(* IEC 61131-3 sources: plc-st-coding-agent/progress/evidence/f14_v6_public_pilot_20261112/jobs/codex_deepseek-v4pro, 32 files *)

(* ---- public-easy-01.candidate_01.st ---- *)
(* ENGINEERING_CONTRACT
Output/Public State | Activation (PUB) | Retention/Hold | Reset/Deactivation (PUB) | Same-Scan Priority | Units/Boundaries
Pump_Motor          | bottleSensor (PUB003) | holds through cleaning | cleaningConfirmButton (PUB004) | stage 0 sensor transition first | BOOL, stages 0..5
Filling_Valve       | cleaningConfirmButton (PUB004) | holds through filling | fillingConfirmButton (PUB005) | current stage only | BOOL
Capping_Machine     | fillingConfirmButton (PUB005) | holds through capping | cappingConfirmButton (PUB006) | current stage only | BOOL
Packing_Machine     | cappingConfirmButton (PUB006) | holds through packing | packingConfirmButton (PUB007) | current stage only | BOOL
Completion_Light    | packingConfirmButton (PUB007) | holds until pickup | finishedButton (PUB008) | stage 5 only | BOOL
Unspecified simultaneous assertions are serialized as one stage transition per scan.
*)
(* CONTRACT_RULES [] *)

FUNCTION_BLOCK AutomatedFillingLine
VAR_INPUT
    bottleSensor : BOOL;
    cleaningConfirmButton : BOOL;
    fillingConfirmButton : BOOL;
    cappingConfirmButton : BOOL;
    packingConfirmButton : BOOL;
    finishedButton : BOOL;
END_VAR
VAR_OUTPUT
    Pump_Motor : BOOL;
    Filling_Valve : BOOL;
    Capping_Machine : BOOL;
    Packing_Machine : BOOL;
    Completion_Light : BOOL;
END_VAR
VAR
    tmp_Stage : INT := 0;
END_VAR

CASE tmp_Stage OF
    0:
        IF bottleSensor THEN
            tmp_Stage := 1;
        END_IF;
    1:
        IF cleaningConfirmButton THEN
            tmp_Stage := 2;
        END_IF;
    2:
        IF fillingConfirmButton THEN
            tmp_Stage := 3;
        END_IF;
    3:
        IF cappingConfirmButton THEN
            tmp_Stage := 4;
        END_IF;
    4:
        IF packingConfirmButton THEN
            tmp_Stage := 5;
        END_IF;
    5:
        IF finishedButton THEN
            tmp_Stage := 0;
        END_IF;
END_CASE;

CASE tmp_Stage OF
    0:
        Pump_Motor := FALSE;
        Filling_Valve := FALSE;
        Capping_Machine := FALSE;
        Packing_Machine := FALSE;
        Completion_Light := FALSE;
    1:
        Pump_Motor := TRUE;
        Filling_Valve := FALSE;
        Capping_Machine := FALSE;
        Packing_Machine := FALSE;
        Completion_Light := FALSE;
    2:
        Pump_Motor := FALSE;
        Filling_Valve := TRUE;
        Capping_Machine := FALSE;
        Packing_Machine := FALSE;
        Completion_Light := FALSE;
    3:
        Pump_Motor := FALSE;
        Filling_Valve := FALSE;
        Capping_Machine := TRUE;
        Packing_Machine := FALSE;
        Completion_Light := FALSE;
    4:
        Pump_Motor := FALSE;
        Filling_Valve := FALSE;
        Capping_Machine := FALSE;
        Packing_Machine := TRUE;
        Completion_Light := FALSE;
    5:
        Pump_Motor := FALSE;
        Filling_Valve := FALSE;
        Capping_Machine := FALSE;
        Packing_Machine := FALSE;
        Completion_Light := TRUE;
END_CASE;

END_FUNCTION_BLOCK

(* ---- public-easy-01.candidate_02.st ---- *)
(* ENGINEERING_CONTRACT
Output/Public State | Activation (PUB) | Retention/Hold | Reset/Deactivation (PUB) | Same-Scan Priority | Units/Boundaries
Pump_Motor          | bottleSensor (PUB003) | holds through entire production cycle | finishedButton (PUB008) | stage 0 sensor transition first | BOOL, stages 0..5
Filling_Valve       | cleaningConfirmButton (PUB004) | holds through filling | fillingConfirmButton (PUB005) | current stage only | BOOL
Capping_Machine     | fillingConfirmButton (PUB005) | holds through capping | cappingConfirmButton (PUB006) | current stage only | BOOL
Packing_Machine     | cappingConfirmButton (PUB006) | holds through packing | packingConfirmButton (PUB007) | current stage only | BOOL
Completion_Light    | packingConfirmButton (PUB007) | holds until pickup | finishedButton (PUB008) | stage 5 only | BOOL
Unspecified simultaneous assertions are serialized as one stage transition per scan.
*)
(* CONTRACT_RULES [] *)

FUNCTION_BLOCK AutomatedFillingLine
VAR_INPUT
    bottleSensor : BOOL;
    cleaningConfirmButton : BOOL;
    fillingConfirmButton : BOOL;
    cappingConfirmButton : BOOL;
    packingConfirmButton : BOOL;
    finishedButton : BOOL;
END_VAR
VAR_OUTPUT
    Pump_Motor : BOOL;
    Filling_Valve : BOOL;
    Capping_Machine : BOOL;
    Packing_Machine : BOOL;
    Completion_Light : BOOL;
END_VAR
VAR
    tmp_Stage : INT := 0;
END_VAR

CASE tmp_Stage OF
    0:
        IF bottleSensor THEN
            tmp_Stage := 1;
        END_IF;
    1:
        IF cleaningConfirmButton THEN
            tmp_Stage := 2;
        END_IF;
    2:
        IF fillingConfirmButton THEN
            tmp_Stage := 3;
        END_IF;
    3:
        IF cappingConfirmButton THEN
            tmp_Stage := 4;
        END_IF;
    4:
        IF packingConfirmButton THEN
            tmp_Stage := 5;
        END_IF;
    5:
        IF finishedButton THEN
            tmp_Stage := 0;
        END_IF;
END_CASE;

CASE tmp_Stage OF
    0:
        Pump_Motor := FALSE;
        Filling_Valve := FALSE;
        Capping_Machine := FALSE;
        Packing_Machine := FALSE;
        Completion_Light := FALSE;
    1:
        Pump_Motor := TRUE;
        Filling_Valve := FALSE;
        Capping_Machine := FALSE;
        Packing_Machine := FALSE;
        Completion_Light := FALSE;
    2:
        Pump_Motor := TRUE;
        Filling_Valve := TRUE;
        Capping_Machine := FALSE;
        Packing_Machine := FALSE;
        Completion_Light := FALSE;
    3:
        Pump_Motor := TRUE;
        Filling_Valve := FALSE;
        Capping_Machine := TRUE;
        Packing_Machine := FALSE;
        Completion_Light := FALSE;
    4:
        Pump_Motor := TRUE;
        Filling_Valve := FALSE;
        Capping_Machine := FALSE;
        Packing_Machine := TRUE;
        Completion_Light := FALSE;
    5:
        Pump_Motor := TRUE;
        Filling_Valve := FALSE;
        Capping_Machine := FALSE;
        Packing_Machine := FALSE;
        Completion_Light := TRUE;
END_CASE;

END_FUNCTION_BLOCK

(* ---- public-easy-01.candidate_03.st ---- *)
(* ENGINEERING_CONTRACT
Output/Public State | Activation (PUB) | Retention/Hold | Reset/Deactivation (PUB) | Same-Scan Priority | Units/Boundaries
Pump_Motor          | bottleSensor (PUB003)         | latched after set through cycle | finishedButton (PUB008) | finishedButton reset wins; then set inputs latch | BOOL
Filling_Valve       | cleaningConfirmButton (PUB004) | latched after set through cycle | finishedButton (PUB008) | finishedButton reset wins; then set inputs latch | BOOL
Capping_Machine     | fillingConfirmButton (PUB005)  | latched after set through cycle | finishedButton (PUB008) | finishedButton reset wins; then set inputs latch | BOOL
Packing_Machine     | cappingConfirmButton (PUB006)  | latched after set through cycle | finishedButton (PUB008) | finishedButton reset wins; then set inputs latch | BOOL
Completion_Light    | packingConfirmButton (PUB007)  | latched after set until pickup | finishedButton (PUB008) | finishedButton reset wins; then set inputs latch | BOOL
All BOOL outputs; no step-enable interlock is applied beyond the specified triggers and finished reset.
*)

(* CONTRACT_RULES [
{"kind":"hold_until_reset","output":"Pump_Motor","set_input":"bottleSensor","reset_input":"finishedButton"},
{"kind":"hold_until_reset","output":"Filling_Valve","set_input":"cleaningConfirmButton","reset_input":"finishedButton"},
{"kind":"hold_until_reset","output":"Capping_Machine","set_input":"fillingConfirmButton","reset_input":"finishedButton"},
{"kind":"hold_until_reset","output":"Packing_Machine","set_input":"cappingConfirmButton","reset_input":"finishedButton"},
{"kind":"hold_until_reset","output":"Completion_Light","set_input":"packingConfirmButton","reset_input":"finishedButton"}
] *)

FUNCTION_BLOCK AutomatedFillingLine
VAR_INPUT
    bottleSensor : BOOL;
    cleaningConfirmButton : BOOL;
    fillingConfirmButton : BOOL;
    cappingConfirmButton : BOOL;
    packingConfirmButton : BOOL;
    finishedButton : BOOL;
END_VAR
VAR_OUTPUT
    Pump_Motor : BOOL;
    Filling_Valve : BOOL;
    Capping_Machine : BOOL;
    Packing_Machine : BOOL;
    Completion_Light : BOOL;
END_VAR

IF finishedButton THEN
    Pump_Motor := FALSE;
    Filling_Valve := FALSE;
    Capping_Machine := FALSE;
    Packing_Machine := FALSE;
    Completion_Light := FALSE;
ELSE
    IF bottleSensor THEN
        Pump_Motor := TRUE;
    END_IF;

    IF cleaningConfirmButton THEN
        Filling_Valve := TRUE;
    END_IF;

    IF fillingConfirmButton THEN
        Capping_Machine := TRUE;
    END_IF;

    IF cappingConfirmButton THEN
        Packing_Machine := TRUE;
    END_IF;

    IF packingConfirmButton THEN
        Completion_Light := TRUE;
    END_IF;
END_IF;

END_FUNCTION_BLOCK

(* ---- public-easy-01.candidate_04.st ---- *)
(* ENGINEERING_CONTRACT
Output/Public State | Activation (PUB) | Retention/Hold | Reset/Deactivation | Same-Scan Priority | Units/Boundaries
Pump_Motor | bottleSensor (PUB003) | latched after cycle start | finishedButton (PUB008) | finished reset wins | BOOL
Filling_Valve | cleaningConfirmButton AND Pump_Motor (PUB004) | latched after start | finishedButton (PUB008) | finished reset wins | BOOL
Capping_Machine | fillingConfirmButton AND Filling_Valve (PUB005) | latched after start | finishedButton (PUB008) | finished reset wins | BOOL
Packing_Machine | cappingConfirmButton AND Capping_Machine (PUB006) | latched after start | finishedButton (PUB008) | finished reset wins | BOOL
Completion_Light | packingConfirmButton AND Packing_Machine (PUB007) | latched until pickup | finishedButton (PUB008) | finished reset wins | BOOL
*)

(* CONTRACT_RULES [
 {"kind":"hold_until_reset","output":"Pump_Motor","set_input":"bottleSensor","reset_input":"finishedButton"}
] *)

FUNCTION_BLOCK AutomatedFillingLine
VAR_INPUT
    bottleSensor : BOOL;
    cleaningConfirmButton : BOOL;
    fillingConfirmButton : BOOL;
    cappingConfirmButton : BOOL;
    packingConfirmButton : BOOL;
    finishedButton : BOOL;
END_VAR
VAR_OUTPUT
    Pump_Motor : BOOL;
    Filling_Valve : BOOL;
    Capping_Machine : BOOL;
    Packing_Machine : BOOL;
    Completion_Light : BOOL;
END_VAR

IF finishedButton THEN
    Pump_Motor := FALSE;
    Filling_Valve := FALSE;
    Capping_Machine := FALSE;
    Packing_Machine := FALSE;
    Completion_Light := FALSE;
ELSE
    IF bottleSensor THEN
        Pump_Motor := TRUE;
    END_IF;

    IF cleaningConfirmButton AND Pump_Motor THEN
        Filling_Valve := TRUE;
    END_IF;

    IF fillingConfirmButton AND Filling_Valve THEN
        Capping_Machine := TRUE;
    END_IF;

    IF cappingConfirmButton AND Capping_Machine THEN
        Packing_Machine := TRUE;
    END_IF;

    IF packingConfirmButton AND Packing_Machine THEN
        Completion_Light := TRUE;
    END_IF;
END_IF;

END_FUNCTION_BLOCK

(* ---- public-easy-01.raw_candidate_01.st ---- *)
(* ENGINEERING_CONTRACT
Output/Public State | Activation (PUB) | Retention/Hold | Reset/Deactivation (PUB) | Same-Scan Priority | Units/Boundaries
Pump_Motor          | bottleSensor (PUB003) | holds through cleaning | cleaningConfirmButton (PUB004) | stage 0 sensor transition first | BOOL, stages 0..5
Filling_Valve       | cleaningConfirmButton (PUB004) | holds through filling | fillingConfirmButton (PUB005) | current stage only | BOOL
Capping_Machine     | fillingConfirmButton (PUB005) | holds through capping | cappingConfirmButton (PUB006) | current stage only | BOOL
Packing_Machine     | cappingConfirmButton (PUB006) | holds through packing | packingConfirmButton (PUB007) | current stage only | BOOL
Completion_Light    | packingConfirmButton (PUB007) | holds until pickup | finishedButton (PUB008) | stage 5 only | BOOL
Unspecified simultaneous assertions are serialized as one stage transition per scan.
*)
(* CONTRACT_RULES [] *)

FUNCTION_BLOCK AutomatedFillingLine
VAR_INPUT
    bottleSensor : BOOL;
    cleaningConfirmButton : BOOL;
    fillingConfirmButton : BOOL;
    cappingConfirmButton : BOOL;
    packingConfirmButton : BOOL;
    finishedButton : BOOL;
END_VAR
VAR_OUTPUT
    Pump_Motor : BOOL;
    Filling_Valve : BOOL;
    Capping_Machine : BOOL;
    Packing_Machine : BOOL;
    Completion_Light : BOOL;
END_VAR
VAR
    tmp_Stage : INT := 0;
END_VAR

CASE tmp_Stage OF
    0:
        IF bottleSensor THEN
            tmp_Stage := 1;
        END_IF;
    1:
        IF cleaningConfirmButton THEN
            tmp_Stage := 2;
        END_IF;
    2:
        IF fillingConfirmButton THEN
            tmp_Stage := 3;
        END_IF;
    3:
        IF cappingConfirmButton THEN
            tmp_Stage := 4;
        END_IF;
    4:
        IF packingConfirmButton THEN
            tmp_Stage := 5;
        END_IF;
    5:
        IF finishedButton THEN
            tmp_Stage := 0;
        END_IF;
END_CASE;

CASE tmp_Stage OF
    0:
        Pump_Motor := FALSE;
        Filling_Valve := FALSE;
        Capping_Machine := FALSE;
        Packing_Machine := FALSE;
        Completion_Light := FALSE;
    1:
        Pump_Motor := TRUE;
        Filling_Valve := FALSE;
        Capping_Machine := FALSE;
        Packing_Machine := FALSE;
        Completion_Light := FALSE;
    2:
        Pump_Motor := FALSE;
        Filling_Valve := TRUE;
        Capping_Machine := FALSE;
        Packing_Machine := FALSE;
        Completion_Light := FALSE;
    3:
        Pump_Motor := FALSE;
        Filling_Valve := FALSE;
        Capping_Machine := TRUE;
        Packing_Machine := FALSE;
        Completion_Light := FALSE;
    4:
        Pump_Motor := FALSE;
        Filling_Valve := FALSE;
        Capping_Machine := FALSE;
        Packing_Machine := TRUE;
        Completion_Light := FALSE;
    5:
        Pump_Motor := FALSE;
        Filling_Valve := FALSE;
        Capping_Machine := FALSE;
        Packing_Machine := FALSE;
        Completion_Light := TRUE;
END_CASE;

END_FUNCTION_BLOCK

(* ---- public-easy-01.raw_candidate_02.st ---- *)
(* ENGINEERING_CONTRACT
Output/Public State | Activation (PUB) | Retention/Hold | Reset/Deactivation (PUB) | Same-Scan Priority | Units/Boundaries
Pump_Motor          | bottleSensor (PUB003) | holds through entire production cycle | finishedButton (PUB008) | stage 0 sensor transition first | BOOL, stages 0..5
Filling_Valve       | cleaningConfirmButton (PUB004) | holds through filling | fillingConfirmButton (PUB005) | current stage only | BOOL
Capping_Machine     | fillingConfirmButton (PUB005) | holds through capping | cappingConfirmButton (PUB006) | current stage only | BOOL
Packing_Machine     | cappingConfirmButton (PUB006) | holds through packing | packingConfirmButton (PUB007) | current stage only | BOOL
Completion_Light    | packingConfirmButton (PUB007) | holds until pickup | finishedButton (PUB008) | stage 5 only | BOOL
Unspecified simultaneous assertions are serialized as one stage transition per scan.
*)
(* CONTRACT_RULES [] *)

FUNCTION_BLOCK AutomatedFillingLine
VAR_INPUT
    bottleSensor : BOOL;
    cleaningConfirmButton : BOOL;
    fillingConfirmButton : BOOL;
    cappingConfirmButton : BOOL;
    packingConfirmButton : BOOL;
    finishedButton : BOOL;
END_VAR
VAR_OUTPUT
    Pump_Motor : BOOL;
    Filling_Valve : BOOL;
    Capping_Machine : BOOL;
    Packing_Machine : BOOL;
    Completion_Light : BOOL;
END_VAR
VAR
    tmp_Stage : INT := 0;
END_VAR

CASE tmp_Stage OF
    0:
        IF bottleSensor THEN
            tmp_Stage := 1;
        END_IF;
    1:
        IF cleaningConfirmButton THEN
            tmp_Stage := 2;
        END_IF;
    2:
        IF fillingConfirmButton THEN
            tmp_Stage := 3;
        END_IF;
    3:
        IF cappingConfirmButton THEN
            tmp_Stage := 4;
        END_IF;
    4:
        IF packingConfirmButton THEN
            tmp_Stage := 5;
        END_IF;
    5:
        IF finishedButton THEN
            tmp_Stage := 0;
        END_IF;
END_CASE;

CASE tmp_Stage OF
    0:
        Pump_Motor := FALSE;
        Filling_Valve := FALSE;
        Capping_Machine := FALSE;
        Packing_Machine := FALSE;
        Completion_Light := FALSE;
    1:
        Pump_Motor := TRUE;
        Filling_Valve := FALSE;
        Capping_Machine := FALSE;
        Packing_Machine := FALSE;
        Completion_Light := FALSE;
    2:
        Pump_Motor := TRUE;
        Filling_Valve := TRUE;
        Capping_Machine := FALSE;
        Packing_Machine := FALSE;
        Completion_Light := FALSE;
    3:
        Pump_Motor := TRUE;
        Filling_Valve := FALSE;
        Capping_Machine := TRUE;
        Packing_Machine := FALSE;
        Completion_Light := FALSE;
    4:
        Pump_Motor := TRUE;
        Filling_Valve := FALSE;
        Capping_Machine := FALSE;
        Packing_Machine := TRUE;
        Completion_Light := FALSE;
    5:
        Pump_Motor := TRUE;
        Filling_Valve := FALSE;
        Capping_Machine := FALSE;
        Packing_Machine := FALSE;
        Completion_Light := TRUE;
END_CASE;

END_FUNCTION_BLOCK

(* ---- public-easy-01.raw_candidate_03.st ---- *)
(* ENGINEERING_CONTRACT
Output/Public State | Activation (PUB) | Retention/Hold | Reset/Deactivation (PUB) | Same-Scan Priority | Units/Boundaries
Pump_Motor          | bottleSensor (PUB003)         | latched after set through cycle | finishedButton (PUB008) | finishedButton reset wins; then set inputs latch | BOOL
Filling_Valve       | cleaningConfirmButton (PUB004) | latched after set through cycle | finishedButton (PUB008) | finishedButton reset wins; then set inputs latch | BOOL
Capping_Machine     | fillingConfirmButton (PUB005)  | latched after set through cycle | finishedButton (PUB008) | finishedButton reset wins; then set inputs latch | BOOL
Packing_Machine     | cappingConfirmButton (PUB006)  | latched after set through cycle | finishedButton (PUB008) | finishedButton reset wins; then set inputs latch | BOOL
Completion_Light    | packingConfirmButton (PUB007)  | latched after set until pickup | finishedButton (PUB008) | finishedButton reset wins; then set inputs latch | BOOL
All BOOL outputs; no step-enable interlock is applied beyond the specified triggers and finished reset.
*)

(* CONTRACT_RULES [
{"kind":"hold_until_reset","output":"Pump_Motor","set_input":"bottleSensor","reset_input":"finishedButton"},
{"kind":"hold_until_reset","output":"Filling_Valve","set_input":"cleaningConfirmButton","reset_input":"finishedButton"},
{"kind":"hold_until_reset","output":"Capping_Machine","set_input":"fillingConfirmButton","reset_input":"finishedButton"},
{"kind":"hold_until_reset","output":"Packing_Machine","set_input":"cappingConfirmButton","reset_input":"finishedButton"},
{"kind":"hold_until_reset","output":"Completion_Light","set_input":"packingConfirmButton","reset_input":"finishedButton"}
] *)

FUNCTION_BLOCK AutomatedFillingLine
VAR_INPUT
    bottleSensor : BOOL;
    cleaningConfirmButton : BOOL;
    fillingConfirmButton : BOOL;
    cappingConfirmButton : BOOL;
    packingConfirmButton : BOOL;
    finishedButton : BOOL;
END_VAR
VAR_OUTPUT
    Pump_Motor : BOOL;
    Filling_Valve : BOOL;
    Capping_Machine : BOOL;
    Packing_Machine : BOOL;
    Completion_Light : BOOL;
END_VAR

IF finishedButton THEN
    Pump_Motor := FALSE;
    Filling_Valve := FALSE;
    Capping_Machine := FALSE;
    Packing_Machine := FALSE;
    Completion_Light := FALSE;
ELSE
    IF bottleSensor THEN
        Pump_Motor := TRUE;
    END_IF;

    IF cleaningConfirmButton THEN
        Filling_Valve := TRUE;
    END_IF;

    IF fillingConfirmButton THEN
        Capping_Machine := TRUE;
    END_IF;

    IF cappingConfirmButton THEN
        Packing_Machine := TRUE;
    END_IF;

    IF packingConfirmButton THEN
        Completion_Light := TRUE;
    END_IF;
END_IF;

END_FUNCTION_BLOCK

(* ---- public-easy-01.raw_candidate_04.st ---- *)
(* ENGINEERING_CONTRACT
Output/Public State | Activation (PUB) | Retention/Hold | Reset/Deactivation | Same-Scan Priority | Units/Boundaries
Pump_Motor | bottleSensor (PUB003) | latched after cycle start | finishedButton (PUB008) | finished reset wins | BOOL
Filling_Valve | cleaningConfirmButton AND Pump_Motor (PUB004) | latched after start | finishedButton (PUB008) | finished reset wins | BOOL
Capping_Machine | fillingConfirmButton AND Filling_Valve (PUB005) | latched after start | finishedButton (PUB008) | finished reset wins | BOOL
Packing_Machine | cappingConfirmButton AND Capping_Machine (PUB006) | latched after start | finishedButton (PUB008) | finished reset wins | BOOL
Completion_Light | packingConfirmButton AND Packing_Machine (PUB007) | latched until pickup | finishedButton (PUB008) | finished reset wins | BOOL
*)

(* CONTRACT_RULES [
 {"kind":"hold_until_reset","output":"Pump_Motor","set_input":"bottleSensor","reset_input":"finishedButton"}
] *)

FUNCTION_BLOCK AutomatedFillingLine
VAR_INPUT
    bottleSensor : BOOL;
    cleaningConfirmButton : BOOL;
    fillingConfirmButton : BOOL;
    cappingConfirmButton : BOOL;
    packingConfirmButton : BOOL;
    finishedButton : BOOL;
END_VAR
VAR_OUTPUT
    Pump_Motor : BOOL;
    Filling_Valve : BOOL;
    Capping_Machine : BOOL;
    Packing_Machine : BOOL;
    Completion_Light : BOOL;
END_VAR

IF finishedButton THEN
    Pump_Motor := FALSE;
    Filling_Valve := FALSE;
    Capping_Machine := FALSE;
    Packing_Machine := FALSE;
    Completion_Light := FALSE;
ELSE
    IF bottleSensor THEN
        Pump_Motor := TRUE;
    END_IF;

    IF cleaningConfirmButton AND Pump_Motor THEN
        Filling_Valve := TRUE;
    END_IF;

    IF fillingConfirmButton AND Filling_Valve THEN
        Capping_Machine := TRUE;
    END_IF;

    IF cappingConfirmButton AND Capping_Machine THEN
        Packing_Machine := TRUE;
    END_IF;

    IF packingConfirmButton AND Packing_Machine THEN
        Completion_Light := TRUE;
    END_IF;
END_IF;

END_FUNCTION_BLOCK

(* ---- public-easy-04.candidate_01.st ---- *)
(*
ENGINEERING_CONTRACT
- VFD_RUN: active iff PASTE_E_STOP_NC AND viscosity_condition; no retention; immediate off on raw FALSE or E_STOP FALSE; PUB003.
- viscosity_condition: becomes TRUE when VISCOSITY_OK TRUE for >= DebounceTime; raw FALSE invalidates immediately; E_STOP clears only incomplete debounce; PUB002/PUB003.
- PUMP_RUNTIME_ACC: adds TIME_TO_LTIME(CycleTime) only when final VFD_RUN TRUE; preserved while stopped; starts at zero; PUB004/PUB006.
- PUMP_MAINT_DUE: TRUE when PUMP_RUNTIME_ACC >= TIME_TO_LTIME(T#500H); informational, no run/permissive effect; PUB005.
- units: DebounceTime/CycleTime TIME ms; accumulated value LTIME ns.
- priority: raw viscosity FALSE and E_STOP FALSE are resolved before same-scan runtime accumulation.
*)
(* CONTRACT_RULES [] *)

FUNCTION_BLOCK JamPumpControl
VAR_INPUT
    VISCOSITY_OK : BOOL;
    PASTE_E_STOP_NC : BOOL;
    DebounceTime : TIME;
    CycleTime : TIME;
END_VAR
VAR_OUTPUT
    VFD_RUN : BOOL;
    PUMP_MAINT_DUE : BOOL;
    PUMP_RUNTIME_ACC : LTIME;
END_VAR
VAR
    local_debounce_elapsed : LTIME := LTIME#0S;
    local_viscosity_condition : BOOL := FALSE;
    local_runtime_accumulator : LTIME := LTIME#0S;
END_VAR

IF VISCOSITY_OK THEN
    IF PASTE_E_STOP_NC THEN
        IF CycleTime > T#0MS THEN
            IF local_debounce_elapsed < TIME_TO_LTIME(DebounceTime) THEN
                local_debounce_elapsed := local_debounce_elapsed + TIME_TO_LTIME(CycleTime);
                IF local_debounce_elapsed > TIME_TO_LTIME(DebounceTime) THEN
                    local_debounce_elapsed := TIME_TO_LTIME(DebounceTime);
                END_IF;
            END_IF;
        END_IF;
    ELSE
        IF local_debounce_elapsed < TIME_TO_LTIME(DebounceTime) THEN
            local_debounce_elapsed := LTIME#0S;
            local_viscosity_condition := FALSE;
        END_IF;
    END_IF;
    local_viscosity_condition := local_debounce_elapsed >= TIME_TO_LTIME(DebounceTime);
ELSE
    local_debounce_elapsed := LTIME#0S;
    local_viscosity_condition := FALSE;
END_IF;

VFD_RUN := PASTE_E_STOP_NC AND local_viscosity_condition;

IF VFD_RUN THEN
    IF CycleTime > T#0MS THEN
        local_runtime_accumulator := local_runtime_accumulator + TIME_TO_LTIME(CycleTime);
    END_IF;
END_IF;

PUMP_RUNTIME_ACC := local_runtime_accumulator;
PUMP_MAINT_DUE := local_runtime_accumulator >= TIME_TO_LTIME(T#500H);

END_FUNCTION_BLOCK

(* ---- public-easy-04.raw_candidate_01.st ---- *)
(*
ENGINEERING_CONTRACT
- VFD_RUN: active iff PASTE_E_STOP_NC AND viscosity_condition; no retention; immediate off on raw FALSE or E_STOP FALSE; PUB003.
- viscosity_condition: becomes TRUE when VISCOSITY_OK TRUE for >= DebounceTime; raw FALSE invalidates immediately; E_STOP clears only incomplete debounce; PUB002/PUB003.
- PUMP_RUNTIME_ACC: adds TIME_TO_LTIME(CycleTime) only when final VFD_RUN TRUE; preserved while stopped; starts at zero; PUB004/PUB006.
- PUMP_MAINT_DUE: TRUE when PUMP_RUNTIME_ACC >= TIME_TO_LTIME(T#500H); informational, no run/permissive effect; PUB005.
- units: DebounceTime/CycleTime TIME ms; accumulated value LTIME ns.
- priority: raw viscosity FALSE and E_STOP FALSE are resolved before same-scan runtime accumulation.
*)
(* CONTRACT_RULES [] *)

FUNCTION_BLOCK JamPumpControl
VAR_INPUT
    VISCOSITY_OK : BOOL;
    PASTE_E_STOP_NC : BOOL;
    DebounceTime : TIME;
    CycleTime : TIME;
END_VAR
VAR_OUTPUT
    VFD_RUN : BOOL;
    PUMP_MAINT_DUE : BOOL;
    PUMP_RUNTIME_ACC : LTIME;
END_VAR
VAR
    local_debounce_elapsed : LTIME := LTIME#0S;
    local_viscosity_condition : BOOL := FALSE;
    local_runtime_accumulator : LTIME := LTIME#0S;
END_VAR

IF VISCOSITY_OK THEN
    IF PASTE_E_STOP_NC THEN
        IF CycleTime > T#0MS THEN
            IF local_debounce_elapsed < TIME_TO_LTIME(DebounceTime) THEN
                local_debounce_elapsed := local_debounce_elapsed + TIME_TO_LTIME(CycleTime);
                IF local_debounce_elapsed > TIME_TO_LTIME(DebounceTime) THEN
                    local_debounce_elapsed := TIME_TO_LTIME(DebounceTime);
                END_IF;
            END_IF;
        END_IF;
    ELSE
        IF local_debounce_elapsed < TIME_TO_LTIME(DebounceTime) THEN
            local_debounce_elapsed := LTIME#0S;
            local_viscosity_condition := FALSE;
        END_IF;
    END_IF;
    local_viscosity_condition := local_debounce_elapsed >= TIME_TO_LTIME(DebounceTime);
ELSE
    local_debounce_elapsed := LTIME#0S;
    local_viscosity_condition := FALSE;
END_IF;

VFD_RUN := PASTE_E_STOP_NC AND local_viscosity_condition;

IF VFD_RUN THEN
    IF CycleTime > T#0MS THEN
        local_runtime_accumulator := local_runtime_accumulator + TIME_TO_LTIME(CycleTime);
    END_IF;
END_IF;

PUMP_RUNTIME_ACC := local_runtime_accumulator;
PUMP_MAINT_DUE := local_runtime_accumulator >= TIME_TO_LTIME(T#500H);

END_FUNCTION_BLOCK

(* ---- public-hard-03.candidate_01.st ---- *)
TYPE ST_Recipe :
STRUCT
    recipeID : INT;
    ingredientType : INT;
    ingredientRatio : REAL;
    productionTemperature : REAL;
END_STRUCT
END_TYPE;

FUNCTION_BLOCK FB_RecipeManager
VAR_INPUT
    addRecipe : BOOL;
    deleteRecipe : BOOL;
    modifyRecipe : BOOL;
    queryRecipe : BOOL;
    recipeIn : ST_Recipe;
END_VAR
VAR_OUTPUT
    recipeAdded : BOOL;
    recipeDeleted : BOOL;
    recipeModified : BOOL;
    recipeQueryResult : ST_Recipe;
    error : BOOL;
    status : WORD;
END_VAR
VAR_IN_OUT
    recipe : ARRAY[1..10] OF ST_Recipe;
END_VAR
VAR
    local_i : INT;
    local_matchIndex : INT;
    local_emptyIndex : INT;
    local_found : BOOL;
    local_emptyFound : BOOL;
    local_activeCommands : INT;
END_VAR

(* ENGINEERING_CONTRACT
  Outputs/database behavior:
  - recipeAdded/recipeDeleted/recipeModified: TRUE only on a successful same-scan command, cleared each scan; no hold.
  - recipeQueryResult: written only on a successful query, cleared at scan start; no retention.
  - error/status: set on command failures per PUB009-PUB012, cleared each scan; no hold.
  - Add order: duplicate=16#8002 before full=16#8003; success fills smallest empty index (PUB010).
  - Delete sets only matching recipeID to 0 (PUB011); modify replaces matching slot (PUB012).
  - recipeID 0 is an empty slot marker. Query/delete/modify of ID 0 returns command-specific failure.
  - Multiple simultaneous commands are unsupported: error=TRUE, status=16#80FF, database unchanged.
  - Bounds: array[1..10], IDs INT, ratios/temperatures REAL (PUB008).
*)

(* CONTRACT_RULES [] *)

recipeAdded := FALSE;
recipeDeleted := FALSE;
recipeModified := FALSE;
recipeQueryResult.recipeID := 0;
recipeQueryResult.ingredientType := 0;
recipeQueryResult.ingredientRatio := 0.0;
recipeQueryResult.productionTemperature := 0.0;
error := FALSE;
status := 16#0000;

local_activeCommands := BOOL_TO_INT(addRecipe) + BOOL_TO_INT(deleteRecipe) + BOOL_TO_INT(modifyRecipe) + BOOL_TO_INT(queryRecipe);

IF local_activeCommands > 1 THEN
    error := TRUE;
    status := 16#80FF;
    RETURN;
END_IF;

IF queryRecipe THEN
    local_found := FALSE;
    local_matchIndex := 0;

    IF recipeIn.recipeID <> 0 THEN
        FOR local_i := 1 TO 10 BY 1 DO
            IF (NOT local_found) AND (recipe[local_i].recipeID = recipeIn.recipeID) THEN
                local_matchIndex := local_i;
                local_found := TRUE;
            END_IF;
        END_FOR;
    END_IF;

    IF local_found THEN
        recipeQueryResult := recipe[local_matchIndex];
        error := FALSE;
        status := 16#0000;
    ELSE
        error := TRUE;
        status := 16#8001;
    END_IF;

ELSIF addRecipe THEN
    local_found := FALSE;
    local_emptyFound := FALSE;
    local_emptyIndex := 0;

    FOR local_i := 1 TO 10 BY 1 DO
        IF recipe[local_i].recipeID = recipeIn.recipeID THEN
            local_found := TRUE;
        END_IF;

        IF (NOT local_emptyFound) AND (recipe[local_i].recipeID = 0) THEN
            local_emptyIndex := local_i;
            local_emptyFound := TRUE;
        END_IF;
    END_FOR;

    IF local_found THEN
        error := TRUE;
        status := 16#8002;
    ELSIF NOT local_emptyFound THEN
        error := TRUE;
        status := 16#8003;
    ELSE
        recipe[local_emptyIndex] := recipeIn;
        recipeAdded := TRUE;
        error := FALSE;
        status := 16#0000;
    END_IF;

ELSIF deleteRecipe THEN
    local_found := FALSE;
    local_matchIndex := 0;

    IF recipeIn.recipeID <> 0 THEN
        FOR local_i := 1 TO 10 BY 1 DO
            IF (NOT local_found) AND (recipe[local_i].recipeID = recipeIn.recipeID) THEN
                local_matchIndex := local_i;
                local_found := TRUE;
            END_IF;
        END_FOR;
    END_IF;

    IF local_found THEN
        recipe[local_matchIndex].recipeID := 0;
        recipeDeleted := TRUE;
        error := FALSE;
        status := 16#0000;
    ELSE
        error := TRUE;
        status := 16#8004;
    END_IF;

ELSIF modifyRecipe THEN
    local_found := FALSE;
    local_matchIndex := 0;

    IF recipeIn.recipeID <> 0 THEN
        FOR local_i := 1 TO 10 BY 1 DO
            IF (NOT local_found) AND (recipe[local_i].recipeID = recipeIn.recipeID) THEN
                local_matchIndex := local_i;
                local_found := TRUE;
            END_IF;
        END_FOR;
    END_IF;

    IF local_found THEN
        recipe[local_matchIndex] := recipeIn;
        recipeModified := TRUE;
        error := FALSE;
        status := 16#0000;
    ELSE
        error := TRUE;
        status := 16#8005;
    END_IF;
END_IF;
END_FUNCTION_BLOCK

(* ---- public-hard-03.candidate_02.st ---- *)
TYPE ST_Recipe :
STRUCT
    recipeID : INT;
    ingredientType : INT;
    ingredientRatio : REAL;
    productionTemperature : REAL;
END_STRUCT
END_TYPE;

FUNCTION_BLOCK FB_RecipeManager
VAR_INPUT
    addRecipe : BOOL;
    deleteRecipe : BOOL;
    modifyRecipe : BOOL;
    queryRecipe : BOOL;
    recipeIn : ST_Recipe;
END_VAR
VAR_OUTPUT
    recipeAdded : BOOL;
    recipeDeleted : BOOL;
    recipeModified : BOOL;
    recipeQueryResult : ST_Recipe;
    error : BOOL;
    status : WORD;
END_VAR
VAR_IN_OUT
    recipe : ARRAY[1..10] OF ST_Recipe;
END_VAR
VAR
    local_i : INT;
    local_matchIndex : INT;
    local_emptyIndex : INT;
    local_found : BOOL;
    local_emptyFound : BOOL;
END_VAR

(* ENGINEERING_CONTRACT
  Outputs/database behavior:
  - recipeAdded/recipeDeleted/recipeModified: pulse TRUE only on a successful same-scan command, cleared at scan start.
  - recipeQueryResult: cleared at scan start; rewritten only on a successful query.
  - error/status: set on command failure per PUB009-PUB012, otherwise no error.
  - Add checks duplicate before full, then stores at smallest empty index (PUB010).
  - Delete clears only the matching recipeID (PUB011); modify replaces the matching slot (PUB012).
  - Query ID not found => error=TRUE, status=16#8001 (PUB009).
  - Add duplicate => 16#8002; add full => 16#8003 (PUB010).
  - Delete ID not found => 16#8004 (PUB011); modify ID not found => 16#8005 (PUB012).
  - recipeID 0 denotes an empty slot (PUB008).
  - Simultaneous commands are unspecified by task text; implemented with interface-order priority:
    addRecipe > deleteRecipe > modifyRecipe > queryRecipe. The higher-priority command is executed,
    lower-priority commands are not processed in that scan.
  - Bounds: ARRAY[1..10], INT and REAL data preserved exactly (PUB008).
*)

(* CONTRACT_RULES [] *)

recipeAdded := FALSE;
recipeDeleted := FALSE;
recipeModified := FALSE;
recipeQueryResult.recipeID := 0;
recipeQueryResult.ingredientType := 0;
recipeQueryResult.ingredientRatio := 0.0;
recipeQueryResult.productionTemperature := 0.0;
error := FALSE;
status := 16#0000;

IF addRecipe THEN
    local_found := FALSE;
    local_emptyFound := FALSE;
    local_emptyIndex := 0;

    FOR local_i := 1 TO 10 BY 1 DO
        IF recipe[local_i].recipeID = recipeIn.recipeID THEN
            local_found := TRUE;
        END_IF;

        IF (NOT local_emptyFound) AND (recipe[local_i].recipeID = 0) THEN
            local_emptyIndex := local_i;
            local_emptyFound := TRUE;
        END_IF;
    END_FOR;

    IF local_found THEN
        error := TRUE;
        status := 16#8002;
    ELSIF NOT local_emptyFound THEN
        error := TRUE;
        status := 16#8003;
    ELSE
        recipe[local_emptyIndex] := recipeIn;
        recipeAdded := TRUE;
        error := FALSE;
        status := 16#0000;
    END_IF;

ELSIF deleteRecipe THEN
    local_found := FALSE;
    local_matchIndex := 0;

    IF recipeIn.recipeID <> 0 THEN
        FOR local_i := 1 TO 10 BY 1 DO
            IF (NOT local_found) AND (recipe[local_i].recipeID = recipeIn.recipeID) THEN
                local_matchIndex := local_i;
                local_found := TRUE;
            END_IF;
        END_FOR;
    END_IF;

    IF local_found THEN
        recipe[local_matchIndex].recipeID := 0;
        recipeDeleted := TRUE;
        error := FALSE;
        status := 16#0000;
    ELSE
        error := TRUE;
        status := 16#8004;
    END_IF;

ELSIF modifyRecipe THEN
    local_found := FALSE;
    local_matchIndex := 0;

    IF recipeIn.recipeID <> 0 THEN
        FOR local_i := 1 TO 10 BY 1 DO
            IF (NOT local_found) AND (recipe[local_i].recipeID = recipeIn.recipeID) THEN
                local_matchIndex := local_i;
                local_found := TRUE;
            END_IF;
        END_FOR;
    END_IF;

    IF local_found THEN
        recipe[local_matchIndex] := recipeIn;
        recipeModified := TRUE;
        error := FALSE;
        status := 16#0000;
    ELSE
        error := TRUE;
        status := 16#8005;
    END_IF;

ELSIF queryRecipe THEN
    local_found := FALSE;
    local_matchIndex := 0;

    IF recipeIn.recipeID <> 0 THEN
        FOR local_i := 1 TO 10 BY 1 DO
            IF (NOT local_found) AND (recipe[local_i].recipeID = recipeIn.recipeID) THEN
                local_matchIndex := local_i;
                local_found := TRUE;
            END_IF;
        END_FOR;
    END_IF;

    IF local_found THEN
        recipeQueryResult := recipe[local_matchIndex];
        error := FALSE;
        status := 16#0000;
    ELSE
        error := TRUE;
        status := 16#8001;
    END_IF;
END_IF;
END_FUNCTION_BLOCK

(* ---- public-hard-03.candidate_03.st ---- *)
TYPE ST_Recipe :
STRUCT
    recipeID : INT;
    ingredientType : INT;
    ingredientRatio : REAL;
    productionTemperature : REAL;
END_STRUCT
END_TYPE;

FUNCTION_BLOCK FB_RecipeManager
VAR_INPUT
    addRecipe : BOOL;
    deleteRecipe : BOOL;
    modifyRecipe : BOOL;
    queryRecipe : BOOL;
    recipeIn : ST_Recipe;
END_VAR
VAR_OUTPUT
    recipeAdded : BOOL;
    recipeDeleted : BOOL;
    recipeModified : BOOL;
    recipeQueryResult : ST_Recipe;
    error : BOOL;
    status : WORD;
END_VAR
VAR_IN_OUT
    recipe : ARRAY[1..10] OF ST_Recipe;
END_VAR
VAR
    local_i : INT;
    local_matchIndex : INT;
    local_emptyIndex : INT;
    local_found : BOOL;
    local_emptyFound : BOOL;
END_VAR

(* ENGINEERING_CONTRACT
  Outputs/database behavior:
  - recipeAdded/recipeDeleted/recipeModified: TRUE only on a successful same-scan command, cleared each scan; no hold.
  - recipeQueryResult: written only on a successful query, cleared at scan start; no retention.
  - error/status: set on command failures per PUB009-PUB012, cleared each scan; no hold.
  - Simultaneous commands: addRecipe has priority; then queryRecipe, deleteRecipe, modifyRecipe.
  - Add order: duplicate=16#8002 before full=16#8003; success fills smallest empty index (PUB010).
  - Delete sets only matching recipeID to 0 (PUB011); modify replaces matching slot (PUB012).
  - recipeID 0 is an empty slot marker. Query/delete/modify of ID 0 returns command-specific failure.
  - Bounds: array[1..10], IDs INT, ratios/temperatures REAL (PUB008).
*)

(* CONTRACT_RULES [] *)

recipeAdded := FALSE;
recipeDeleted := FALSE;
recipeModified := FALSE;
recipeQueryResult.recipeID := 0;
recipeQueryResult.ingredientType := 0;
recipeQueryResult.ingredientRatio := 0.0;
recipeQueryResult.productionTemperature := 0.0;
error := FALSE;
status := 16#0000;

IF addRecipe THEN
    local_found := FALSE;
    local_emptyFound := FALSE;
    local_emptyIndex := 0;

    FOR local_i := 1 TO 10 BY 1 DO
        IF recipe[local_i].recipeID = recipeIn.recipeID THEN
            local_found := TRUE;
        END_IF;

        IF (NOT local_emptyFound) AND (recipe[local_i].recipeID = 0) THEN
            local_emptyIndex := local_i;
            local_emptyFound := TRUE;
        END_IF;
    END_FOR;

    IF local_found THEN
        error := TRUE;
        status := 16#8002;
    ELSIF NOT local_emptyFound THEN
        error := TRUE;
        status := 16#8003;
    ELSE
        recipe[local_emptyIndex] := recipeIn;
        recipeAdded := TRUE;
        error := FALSE;
        status := 16#0000;
    END_IF;

ELSIF queryRecipe THEN
    local_found := FALSE;
    local_matchIndex := 0;

    IF recipeIn.recipeID <> 0 THEN
        FOR local_i := 1 TO 10 BY 1 DO
            IF (NOT local_found) AND (recipe[local_i].recipeID = recipeIn.recipeID) THEN
                local_matchIndex := local_i;
                local_found := TRUE;
            END_IF;
        END_FOR;
    END_IF;

    IF local_found THEN
        recipeQueryResult := recipe[local_matchIndex];
        error := FALSE;
        status := 16#0000;
    ELSE
        error := TRUE;
        status := 16#8001;
    END_IF;

ELSIF deleteRecipe THEN
    local_found := FALSE;
    local_matchIndex := 0;

    IF recipeIn.recipeID <> 0 THEN
        FOR local_i := 1 TO 10 BY 1 DO
            IF (NOT local_found) AND (recipe[local_i].recipeID = recipeIn.recipeID) THEN
                local_matchIndex := local_i;
                local_found := TRUE;
            END_IF;
        END_FOR;
    END_IF;

    IF local_found THEN
        recipe[local_matchIndex].recipeID := 0;
        recipeDeleted := TRUE;
        error := FALSE;
        status := 16#0000;
    ELSE
        error := TRUE;
        status := 16#8004;
    END_IF;

ELSIF modifyRecipe THEN
    local_found := FALSE;
    local_matchIndex := 0;

    IF recipeIn.recipeID <> 0 THEN
        FOR local_i := 1 TO 10 BY 1 DO
            IF (NOT local_found) AND (recipe[local_i].recipeID = recipeIn.recipeID) THEN
                local_matchIndex := local_i;
                local_found := TRUE;
            END_IF;
        END_FOR;
    END_IF;

    IF local_found THEN
        recipe[local_matchIndex] := recipeIn;
        recipeModified := TRUE;
        error := FALSE;
        status := 16#0000;
    ELSE
        error := TRUE;
        status := 16#8005;
    END_IF;
END_IF;
END_FUNCTION_BLOCK

(* ---- public-hard-03.candidate_04.st ---- *)
TYPE ST_Recipe :
STRUCT
    recipeID : INT;
    ingredientType : INT;
    ingredientRatio : REAL;
    productionTemperature : REAL;
END_STRUCT
END_TYPE;

FUNCTION_BLOCK FB_RecipeManager
VAR_INPUT
    addRecipe : BOOL;
    deleteRecipe : BOOL;
    modifyRecipe : BOOL;
    queryRecipe : BOOL;
    recipeIn : ST_Recipe;
END_VAR
VAR_OUTPUT
    recipeAdded : BOOL;
    recipeDeleted : BOOL;
    recipeModified : BOOL;
    recipeQueryResult : ST_Recipe;
    error : BOOL;
    status : WORD;
END_VAR
VAR_IN_OUT
    recipe : ARRAY[1..10] OF ST_Recipe;
END_VAR
VAR
    local_i : INT;
    local_matchIndex : INT;
    local_emptyIndex : INT;
    local_found : BOOL;
    local_emptyFound : BOOL;
END_VAR

(* ENGINEERING_CONTRACT
  Outputs/database behavior:
  - recipeAdded/recipeDeleted/recipeModified: TRUE only on a successful same-scan command, cleared each scan; no hold.
  - recipeQueryResult: written only on a successful query, cleared at scan start; no retention.
  - error/status: set on command failures per PUB009-PUB012, cleared each scan; no hold.
  - Add order: duplicate=16#8002 before full=16#8003; success fills smallest empty index (PUB010).
  - Delete sets only matching recipeID to 0 (PUB011); modify replaces matching slot (PUB012).
  - recipeID 0 is an empty slot marker. Query/delete/modify of ID 0 returns command-specific failure.
  - Multiple simultaneous commands are unspecified by PUB. Consistent interpretation: add > delete > modify > query.
  - Bounds: array[1..10], IDs INT, ratios/temperatures REAL (PUB008).
*)

(* CONTRACT_RULES [] *)

recipeAdded := FALSE;
recipeDeleted := FALSE;
recipeModified := FALSE;
recipeQueryResult.recipeID := 0;
recipeQueryResult.ingredientType := 0;
recipeQueryResult.ingredientRatio := 0.0;
recipeQueryResult.productionTemperature := 0.0;
error := FALSE;
status := 16#0000;

IF addRecipe THEN
    local_found := FALSE;
    local_emptyFound := FALSE;
    local_emptyIndex := 0;

    FOR local_i := 1 TO 10 BY 1 DO
        IF recipe[local_i].recipeID = recipeIn.recipeID THEN
            local_found := TRUE;
        END_IF;

        IF (NOT local_emptyFound) AND (recipe[local_i].recipeID = 0) THEN
            local_emptyIndex := local_i;
            local_emptyFound := TRUE;
        END_IF;
    END_FOR;

    IF local_found THEN
        error := TRUE;
        status := 16#8002;
    ELSIF NOT local_emptyFound THEN
        error := TRUE;
        status := 16#8003;
    ELSE
        recipe[local_emptyIndex] := recipeIn;
        recipeAdded := TRUE;
        error := FALSE;
        status := 16#0000;
    END_IF;

ELSIF deleteRecipe THEN
    local_found := FALSE;
    local_matchIndex := 0;

    IF recipeIn.recipeID <> 0 THEN
        FOR local_i := 1 TO 10 BY 1 DO
            IF (NOT local_found) AND (recipe[local_i].recipeID = recipeIn.recipeID) THEN
                local_matchIndex := local_i;
                local_found := TRUE;
            END_IF;
        END_FOR;
    END_IF;

    IF local_found THEN
        recipe[local_matchIndex].recipeID := 0;
        recipeDeleted := TRUE;
        error := FALSE;
        status := 16#0000;
    ELSE
        error := TRUE;
        status := 16#8004;
    END_IF;

ELSIF modifyRecipe THEN
    local_found := FALSE;
    local_matchIndex := 0;

    IF recipeIn.recipeID <> 0 THEN
        FOR local_i := 1 TO 10 BY 1 DO
            IF (NOT local_found) AND (recipe[local_i].recipeID = recipeIn.recipeID) THEN
                local_matchIndex := local_i;
                local_found := TRUE;
            END_IF;
        END_FOR;
    END_IF;

    IF local_found THEN
        recipe[local_matchIndex] := recipeIn;
        recipeModified := TRUE;
        error := FALSE;
        status := 16#0000;
    ELSE
        error := TRUE;
        status := 16#8005;
    END_IF;

ELSIF queryRecipe THEN
    local_found := FALSE;
    local_matchIndex := 0;

    IF recipeIn.recipeID <> 0 THEN
        FOR local_i := 1 TO 10 BY 1 DO
            IF (NOT local_found) AND (recipe[local_i].recipeID = recipeIn.recipeID) THEN
                local_matchIndex := local_i;
                local_found := TRUE;
            END_IF;
        END_FOR;
    END_IF;

    IF local_found THEN
        recipeQueryResult := recipe[local_matchIndex];
        error := FALSE;
        status := 16#0000;
    ELSE
        error := TRUE;
        status := 16#8001;
    END_IF;
END_IF;

END_FUNCTION_BLOCK

(* ---- public-hard-03.raw_candidate_01.st ---- *)
TYPE ST_Recipe :
STRUCT
    recipeID : INT;
    ingredientType : INT;
    ingredientRatio : REAL;
    productionTemperature : REAL;
END_STRUCT
END_TYPE

FUNCTION_BLOCK FB_RecipeManager
VAR_INPUT
    addRecipe : BOOL;
    deleteRecipe : BOOL;
    modifyRecipe : BOOL;
    queryRecipe : BOOL;
    recipeIn : ST_Recipe;
END_VAR
VAR_OUTPUT
    recipeAdded : BOOL;
    recipeDeleted : BOOL;
    recipeModified : BOOL;
    recipeQueryResult : ST_Recipe;
    error : BOOL;
    status : WORD;
END_VAR
VAR_IN_OUT
    recipe : ARRAY[1..10] OF ST_Recipe;
END_VAR
VAR
    local_i : INT;
    local_matchIndex : INT;
    local_emptyIndex : INT;
    local_found : BOOL;
    local_emptyFound : BOOL;
    local_activeCommands : INT;
END_VAR

(* ENGINEERING_CONTRACT
  Outputs/database behavior:
  - recipeAdded/recipeDeleted/recipeModified: TRUE only on a successful same-scan command, cleared each scan; no hold.
  - recipeQueryResult: written only on a successful query, cleared at scan start; no retention.
  - error/status: set on command failures per PUB009-PUB012, cleared each scan; no hold.
  - Add order: duplicate=16#8002 before full=16#8003; success fills smallest empty index (PUB010).
  - Delete sets only matching recipeID to 0 (PUB011); modify replaces matching slot (PUB012).
  - recipeID 0 is an empty slot marker. Query/delete/modify of ID 0 returns command-specific failure.
  - Multiple simultaneous commands are unsupported: error=TRUE, status=16#80FF, database unchanged.
  - Bounds: array[1..10], IDs INT, ratios/temperatures REAL (PUB008).
*)

(* CONTRACT_RULES [] *)

recipeAdded := FALSE;
recipeDeleted := FALSE;
recipeModified := FALSE;
recipeQueryResult.recipeID := 0;
recipeQueryResult.ingredientType := 0;
recipeQueryResult.ingredientRatio := 0.0;
recipeQueryResult.productionTemperature := 0.0;
error := FALSE;
status := 16#0000;

local_activeCommands := BOOL_TO_INT(addRecipe) + BOOL_TO_INT(deleteRecipe) + BOOL_TO_INT(modifyRecipe) + BOOL_TO_INT(queryRecipe);

IF local_activeCommands > 1 THEN
    error := TRUE;
    status := 16#80FF;
    RETURN;
END_IF;

IF queryRecipe THEN
    local_found := FALSE;
    local_matchIndex := 0;

    IF recipeIn.recipeID <> 0 THEN
        FOR local_i := 1 TO 10 BY 1 DO
            IF (NOT local_found) AND (recipe[local_i].recipeID = recipeIn.recipeID) THEN
                local_matchIndex := local_i;
                local_found := TRUE;
            END_IF;
        END_FOR;
    END_IF;

    IF local_found THEN
        recipeQueryResult := recipe[local_matchIndex];
        error := FALSE;
        status := 16#0000;
    ELSE
        error := TRUE;
        status := 16#8001;
    END_IF;

ELSIF addRecipe THEN
    local_found := FALSE;
    local_emptyFound := FALSE;
    local_emptyIndex := 0;

    FOR local_i := 1 TO 10 BY 1 DO
        IF recipe[local_i].recipeID = recipeIn.recipeID THEN
            local_found := TRUE;
        END_IF;

        IF (NOT local_emptyFound) AND (recipe[local_i].recipeID = 0) THEN
            local_emptyIndex := local_i;
            local_emptyFound := TRUE;
        END_IF;
    END_FOR;

    IF local_found THEN
        error := TRUE;
        status := 16#8002;
    ELSIF NOT local_emptyFound THEN
        error := TRUE;
        status := 16#8003;
    ELSE
        recipe[local_emptyIndex] := recipeIn;
        recipeAdded := TRUE;
        error := FALSE;
        status := 16#0000;
    END_IF;

ELSIF deleteRecipe THEN
    local_found := FALSE;
    local_matchIndex := 0;

    IF recipeIn.recipeID <> 0 THEN
        FOR local_i := 1 TO 10 BY 1 DO
            IF (NOT local_found) AND (recipe[local_i].recipeID = recipeIn.recipeID) THEN
                local_matchIndex := local_i;
                local_found := TRUE;
            END_IF;
        END_FOR;
    END_IF;

    IF local_found THEN
        recipe[local_matchIndex].recipeID := 0;
        recipeDeleted := TRUE;
        error := FALSE;
        status := 16#0000;
    ELSE
        error := TRUE;
        status := 16#8004;
    END_IF;

ELSIF modifyRecipe THEN
    local_found := FALSE;
    local_matchIndex := 0;

    IF recipeIn.recipeID <> 0 THEN
        FOR local_i := 1 TO 10 BY 1 DO
            IF (NOT local_found) AND (recipe[local_i].recipeID = recipeIn.recipeID) THEN
                local_matchIndex := local_i;
                local_found := TRUE;
            END_IF;
        END_FOR;
    END_IF;

    IF local_found THEN
        recipe[local_matchIndex] := recipeIn;
        recipeModified := TRUE;
        error := FALSE;
        status := 16#0000;
    ELSE
        error := TRUE;
        status := 16#8005;
    END_IF;
END_IF;
END_FUNCTION_BLOCK

(* ---- public-hard-03.raw_candidate_02.st ---- *)
TYPE ST_Recipe :
STRUCT
    recipeID : INT;
    ingredientType : INT;
    ingredientRatio : REAL;
    productionTemperature : REAL;
END_STRUCT
END_TYPE;

FUNCTION_BLOCK FB_RecipeManager
VAR_INPUT
    addRecipe : BOOL;
    deleteRecipe : BOOL;
    modifyRecipe : BOOL;
    queryRecipe : BOOL;
    recipeIn : ST_Recipe;
END_VAR
VAR_OUTPUT
    recipeAdded : BOOL;
    recipeDeleted : BOOL;
    recipeModified : BOOL;
    recipeQueryResult : ST_Recipe;
    error : BOOL;
    status : WORD;
END_VAR
VAR_IN_OUT
    recipe : ARRAY[1..10] OF ST_Recipe;
END_VAR
VAR
    local_i : INT;
    local_matchIndex : INT;
    local_emptyIndex : INT;
    local_found : BOOL;
    local_emptyFound : BOOL;
END_VAR

(* ENGINEERING_CONTRACT
  Outputs/database behavior:
  - recipeAdded/recipeDeleted/recipeModified: pulse TRUE only on a successful same-scan command, cleared at scan start.
  - recipeQueryResult: cleared at scan start; rewritten only on a successful query.
  - error/status: set on command failure per PUB009-PUB012, otherwise no error.
  - Add checks duplicate before full, then stores at smallest empty index (PUB010).
  - Delete clears only the matching recipeID (PUB011); modify replaces the matching slot (PUB012).
  - Query ID not found => error=TRUE, status=16#8001 (PUB009).
  - Add duplicate => 16#8002; add full => 16#8003 (PUB010).
  - Delete ID not found => 16#8004 (PUB011); modify ID not found => 16#8005 (PUB012).
  - recipeID 0 denotes an empty slot (PUB008).
  - Simultaneous commands are unspecified by task text; implemented with interface-order priority:
    addRecipe > deleteRecipe > modifyRecipe > queryRecipe. The higher-priority command is executed,
    lower-priority commands are not processed in that scan.
  - Bounds: ARRAY[1..10], INT and REAL data preserved exactly (PUB008).
*)

(* CONTRACT_RULES [] *)

recipeAdded := FALSE;
recipeDeleted := FALSE;
recipeModified := FALSE;
recipeQueryResult.recipeID := 0;
recipeQueryResult.ingredientType := 0;
recipeQueryResult.ingredientRatio := 0.0;
recipeQueryResult.productionTemperature := 0.0;
error := FALSE;
status := 16#0000;

IF addRecipe THEN
    local_found := FALSE;
    local_emptyFound := FALSE;
    local_emptyIndex := 0;

    FOR local_i := 1 TO 10 BY 1 DO
        IF recipe[local_i].recipeID = recipeIn.recipeID THEN
            local_found := TRUE;
        END_IF;

        IF (NOT local_emptyFound) AND (recipe[local_i].recipeID = 0) THEN
            local_emptyIndex := local_i;
            local_emptyFound := TRUE;
        END_IF;
    END_FOR;

    IF local_found THEN
        error := TRUE;
        status := 16#8002;
    ELSIF NOT local_emptyFound THEN
        error := TRUE;
        status := 16#8003;
    ELSE
        recipe[local_emptyIndex] := recipeIn;
        recipeAdded := TRUE;
        error := FALSE;
        status := 16#0000;
    END_IF;

ELSIF deleteRecipe THEN
    local_found := FALSE;
    local_matchIndex := 0;

    IF recipeIn.recipeID <> 0 THEN
        FOR local_i := 1 TO 10 BY 1 DO
            IF (NOT local_found) AND (recipe[local_i].recipeID = recipeIn.recipeID) THEN
                local_matchIndex := local_i;
                local_found := TRUE;
            END_IF;
        END_FOR;
    END_IF;

    IF local_found THEN
        recipe[local_matchIndex].recipeID := 0;
        recipeDeleted := TRUE;
        error := FALSE;
        status := 16#0000;
    ELSE
        error := TRUE;
        status := 16#8004;
    END_IF;

ELSIF modifyRecipe THEN
    local_found := FALSE;
    local_matchIndex := 0;

    IF recipeIn.recipeID <> 0 THEN
        FOR local_i := 1 TO 10 BY 1 DO
            IF (NOT local_found) AND (recipe[local_i].recipeID = recipeIn.recipeID) THEN
                local_matchIndex := local_i;
                local_found := TRUE;
            END_IF;
        END_FOR;
    END_IF;

    IF local_found THEN
        recipe[local_matchIndex] := recipeIn;
        recipeModified := TRUE;
        error := FALSE;
        status := 16#0000;
    ELSE
        error := TRUE;
        status := 16#8005;
    END_IF;

ELSIF queryRecipe THEN
    local_found := FALSE;
    local_matchIndex := 0;

    IF recipeIn.recipeID <> 0 THEN
        FOR local_i := 1 TO 10 BY 1 DO
            IF (NOT local_found) AND (recipe[local_i].recipeID = recipeIn.recipeID) THEN
                local_matchIndex := local_i;
                local_found := TRUE;
            END_IF;
        END_FOR;
    END_IF;

    IF local_found THEN
        recipeQueryResult := recipe[local_matchIndex];
        error := FALSE;
        status := 16#0000;
    ELSE
        error := TRUE;
        status := 16#8001;
    END_IF;
END_IF;
END_FUNCTION_BLOCK

(* ---- public-hard-03.raw_candidate_03.st ---- *)
TYPE ST_Recipe :
STRUCT
    recipeID : INT;
    ingredientType : INT;
    ingredientRatio : REAL;
    productionTemperature : REAL;
END_STRUCT
END_TYPE;

FUNCTION_BLOCK FB_RecipeManager
VAR_INPUT
    addRecipe : BOOL;
    deleteRecipe : BOOL;
    modifyRecipe : BOOL;
    queryRecipe : BOOL;
    recipeIn : ST_Recipe;
END_VAR
VAR_OUTPUT
    recipeAdded : BOOL;
    recipeDeleted : BOOL;
    recipeModified : BOOL;
    recipeQueryResult : ST_Recipe;
    error : BOOL;
    status : WORD;
END_VAR
VAR_IN_OUT
    recipe : ARRAY[1..10] OF ST_Recipe;
END_VAR
VAR
    local_i : INT;
    local_matchIndex : INT;
    local_emptyIndex : INT;
    local_found : BOOL;
    local_emptyFound : BOOL;
END_VAR

(* ENGINEERING_CONTRACT
  Outputs/database behavior:
  - recipeAdded/recipeDeleted/recipeModified: TRUE only on a successful same-scan command, cleared each scan; no hold.
  - recipeQueryResult: written only on a successful query, cleared at scan start; no retention.
  - error/status: set on command failures per PUB009-PUB012, cleared each scan; no hold.
  - Simultaneous commands: addRecipe has priority; then queryRecipe, deleteRecipe, modifyRecipe.
  - Add order: duplicate=16#8002 before full=16#8003; success fills smallest empty index (PUB010).
  - Delete sets only matching recipeID to 0 (PUB011); modify replaces matching slot (PUB012).
  - recipeID 0 is an empty slot marker. Query/delete/modify of ID 0 returns command-specific failure.
  - Bounds: array[1..10], IDs INT, ratios/temperatures REAL (PUB008).
*)

(* CONTRACT_RULES [] *)

recipeAdded := FALSE;
recipeDeleted := FALSE;
recipeModified := FALSE;
recipeQueryResult.recipeID := 0;
recipeQueryResult.ingredientType := 0;
recipeQueryResult.ingredientRatio := 0.0;
recipeQueryResult.productionTemperature := 0.0;
error := FALSE;
status := 16#0000;

IF addRecipe THEN
    local_found := FALSE;
    local_emptyFound := FALSE;
    local_emptyIndex := 0;

    FOR local_i := 1 TO 10 BY 1 DO
        IF recipe[local_i].recipeID = recipeIn.recipeID THEN
            local_found := TRUE;
        END_IF;

        IF (NOT local_emptyFound) AND (recipe[local_i].recipeID = 0) THEN
            local_emptyIndex := local_i;
            local_emptyFound := TRUE;
        END_IF;
    END_FOR;

    IF local_found THEN
        error := TRUE;
        status := 16#8002;
    ELSIF NOT local_emptyFound THEN
        error := TRUE;
        status := 16#8003;
    ELSE
        recipe[local_emptyIndex] := recipeIn;
        recipeAdded := TRUE;
        error := FALSE;
        status := 16#0000;
    END_IF;

ELSIF queryRecipe THEN
    local_found := FALSE;
    local_matchIndex := 0;

    IF recipeIn.recipeID <> 0 THEN
        FOR local_i := 1 TO 10 BY 1 DO
            IF (NOT local_found) AND (recipe[local_i].recipeID = recipeIn.recipeID) THEN
                local_matchIndex := local_i;
                local_found := TRUE;
            END_IF;
        END_FOR;
    END_IF;

    IF local_found THEN
        recipeQueryResult := recipe[local_matchIndex];
        error := FALSE;
        status := 16#0000;
    ELSE
        error := TRUE;
        status := 16#8001;
    END_IF;

ELSIF deleteRecipe THEN
    local_found := FALSE;
    local_matchIndex := 0;

    IF recipeIn.recipeID <> 0 THEN
        FOR local_i := 1 TO 10 BY 1 DO
            IF (NOT local_found) AND (recipe[local_i].recipeID = recipeIn.recipeID) THEN
                local_matchIndex := local_i;
                local_found := TRUE;
            END_IF;
        END_FOR;
    END_IF;

    IF local_found THEN
        recipe[local_matchIndex].recipeID := 0;
        recipeDeleted := TRUE;
        error := FALSE;
        status := 16#0000;
    ELSE
        error := TRUE;
        status := 16#8004;
    END_IF;

ELSIF modifyRecipe THEN
    local_found := FALSE;
    local_matchIndex := 0;

    IF recipeIn.recipeID <> 0 THEN
        FOR local_i := 1 TO 10 BY 1 DO
            IF (NOT local_found) AND (recipe[local_i].recipeID = recipeIn.recipeID) THEN
                local_matchIndex := local_i;
                local_found := TRUE;
            END_IF;
        END_FOR;
    END_IF;

    IF local_found THEN
        recipe[local_matchIndex] := recipeIn;
        recipeModified := TRUE;
        error := FALSE;
        status := 16#0000;
    ELSE
        error := TRUE;
        status := 16#8005;
    END_IF;
END_IF;
END_FUNCTION_BLOCK

(* ---- public-hard-03.raw_candidate_04.st ---- *)
TYPE ST_Recipe :
STRUCT
    recipeID : INT;
    ingredientType : INT;
    ingredientRatio : REAL;
    productionTemperature : REAL;
END_STRUCT
END_TYPE;

FUNCTION_BLOCK FB_RecipeManager
VAR_INPUT
    addRecipe : BOOL;
    deleteRecipe : BOOL;
    modifyRecipe : BOOL;
    queryRecipe : BOOL;
    recipeIn : ST_Recipe;
END_VAR
VAR_OUTPUT
    recipeAdded : BOOL;
    recipeDeleted : BOOL;
    recipeModified : BOOL;
    recipeQueryResult : ST_Recipe;
    error : BOOL;
    status : WORD;
END_VAR
VAR_IN_OUT
    recipe : ARRAY[1..10] OF ST_Recipe;
END_VAR
VAR
    local_i : INT;
    local_matchIndex : INT;
    local_emptyIndex : INT;
    local_found : BOOL;
    local_emptyFound : BOOL;
END_VAR

(* ENGINEERING_CONTRACT
  Outputs/database behavior:
  - recipeAdded/recipeDeleted/recipeModified: TRUE only on a successful same-scan command, cleared each scan; no hold.
  - recipeQueryResult: written only on a successful query, cleared at scan start; no retention.
  - error/status: set on command failures per PUB009-PUB012, cleared each scan; no hold.
  - Add order: duplicate=16#8002 before full=16#8003; success fills smallest empty index (PUB010).
  - Delete sets only matching recipeID to 0 (PUB011); modify replaces matching slot (PUB012).
  - recipeID 0 is an empty slot marker. Query/delete/modify of ID 0 returns command-specific failure.
  - Multiple simultaneous commands are unspecified by PUB. Consistent interpretation: add > delete > modify > query.
  - Bounds: array[1..10], IDs INT, ratios/temperatures REAL (PUB008).
*)

(* CONTRACT_RULES [] *)

recipeAdded := FALSE;
recipeDeleted := FALSE;
recipeModified := FALSE;
recipeQueryResult.recipeID := 0;
recipeQueryResult.ingredientType := 0;
recipeQueryResult.ingredientRatio := 0.0;
recipeQueryResult.productionTemperature := 0.0;
error := FALSE;
status := 16#0000;

IF addRecipe THEN
    local_found := FALSE;
    local_emptyFound := FALSE;
    local_emptyIndex := 0;

    FOR local_i := 1 TO 10 BY 1 DO
        IF recipe[local_i].recipeID = recipeIn.recipeID THEN
            local_found := TRUE;
        END_IF;

        IF (NOT local_emptyFound) AND (recipe[local_i].recipeID = 0) THEN
            local_emptyIndex := local_i;
            local_emptyFound := TRUE;
        END_IF;
    END_FOR;

    IF local_found THEN
        error := TRUE;
        status := 16#8002;
    ELSIF NOT local_emptyFound THEN
        error := TRUE;
        status := 16#8003;
    ELSE
        recipe[local_emptyIndex] := recipeIn;
        recipeAdded := TRUE;
        error := FALSE;
        status := 16#0000;
    END_IF;

ELSIF deleteRecipe THEN
    local_found := FALSE;
    local_matchIndex := 0;

    IF recipeIn.recipeID <> 0 THEN
        FOR local_i := 1 TO 10 BY 1 DO
            IF (NOT local_found) AND (recipe[local_i].recipeID = recipeIn.recipeID) THEN
                local_matchIndex := local_i;
                local_found := TRUE;
            END_IF;
        END_FOR;
    END_IF;

    IF local_found THEN
        recipe[local_matchIndex].recipeID := 0;
        recipeDeleted := TRUE;
        error := FALSE;
        status := 16#0000;
    ELSE
        error := TRUE;
        status := 16#8004;
    END_IF;

ELSIF modifyRecipe THEN
    local_found := FALSE;
    local_matchIndex := 0;

    IF recipeIn.recipeID <> 0 THEN
        FOR local_i := 1 TO 10 BY 1 DO
            IF (NOT local_found) AND (recipe[local_i].recipeID = recipeIn.recipeID) THEN
                local_matchIndex := local_i;
                local_found := TRUE;
            END_IF;
        END_FOR;
    END_IF;

    IF local_found THEN
        recipe[local_matchIndex] := recipeIn;
        recipeModified := TRUE;
        error := FALSE;
        status := 16#0000;
    ELSE
        error := TRUE;
        status := 16#8005;
    END_IF;

ELSIF queryRecipe THEN
    local_found := FALSE;
    local_matchIndex := 0;

    IF recipeIn.recipeID <> 0 THEN
        FOR local_i := 1 TO 10 BY 1 DO
            IF (NOT local_found) AND (recipe[local_i].recipeID = recipeIn.recipeID) THEN
                local_matchIndex := local_i;
                local_found := TRUE;
            END_IF;
        END_FOR;
    END_IF;

    IF local_found THEN
        recipeQueryResult := recipe[local_matchIndex];
        error := FALSE;
        status := 16#0000;
    ELSE
        error := TRUE;
        status := 16#8001;
    END_IF;
END_IF;

END_FUNCTION_BLOCK

(* ---- public-medium-03.candidate_01.st ---- *)
(* ENGINEERING_CONTRACT
average: activated when a sample is accepted; otherwise holds last valid result; reset sets it to 0.0; units are inherited from value (LREAL).
windowSizeReached: TRUE when accepted sample count >= windowSize; holds until reset or invalid window; no edge-only behavior.
error/status: windowSize < 1 or windowSize > 100 sets error=TRUE and status=16#8200; valid window sets error=FALSE and status=16#0000.
capture priority: cyclicExecution=TRUE captures every scan and suppresses trigger; trigger uses R_TRIG only while cyclicExecution=FALSE; reset suppresses capture.
reset: level-triggered on reset=TRUE, clears sum, buffer count, write index, average, and windowSizeReached.
invalid window preserves accumulated average data but forces windowSizeReached=FALSE and prevents new samples.
Boundaries: windowSize is 1..100; storage is ARRAY[0..99] OF LREAL; average division uses INT_TO_LREAL.
PUB001, PUB002, PUB003, PUB004, PUB006, PUB007.
*)
(* CONTRACT_RULES [] *)

FUNCTION_BLOCK FB
VAR_INPUT
    cyclicExecution : BOOL;
    trigger : BOOL;
    value : LREAL;
    windowSize : INT;
    reset : BOOL;
END_VAR
VAR_OUTPUT
    average : LREAL;
    windowSizeReached : BOOL;
    error : BOOL;
    status : WORD;
END_VAR
VAR
    local_buffer : ARRAY[0..99] OF LREAL;
    local_count : INT;
    local_write_index : INT;
    local_sum : LREAL;
    local_trigger_rt : R_TRIG;
END_VAR

local_trigger_rt(CLK := trigger);

IF reset THEN
    local_count := 0;
    local_write_index := 0;
    local_sum := 0.0;
    average := 0.0;
    windowSizeReached := FALSE;
END_IF;

IF (windowSize < 1) OR (windowSize > 100) THEN
    error := TRUE;
    status := 16#8200;
    windowSizeReached := FALSE;
ELSE
    error := FALSE;
    status := 16#0000;

    IF NOT reset THEN
        IF cyclicExecution OR (local_trigger_rt.Q AND (NOT cyclicExecution)) THEN
            IF local_count < windowSize THEN
                local_buffer[local_count] := value;
                local_sum := local_sum + value;
                local_count := local_count + 1;
            ELSE
                local_sum := local_sum - local_buffer[local_write_index] + value;
                local_buffer[local_write_index] := value;
                local_write_index := local_write_index + 1;
                IF local_write_index >= windowSize THEN
                    local_write_index := 0;
                END_IF;
            END_IF;

            IF local_count > 0 THEN
                average := local_sum / INT_TO_LREAL(local_count);
            END_IF;

            windowSizeReached := local_count >= windowSize;
        END_IF;
    END_IF;
END_IF;

END_FUNCTION_BLOCK

(* ---- public-medium-03.candidate_02.st ---- *)
(* ENGINEERING_CONTRACT
average: updates on each accepted sample (PUB002/PUB003), holds between samples; reset=TRUE clears it in the same scan; units LREAL.
windowSizeReached: TRUE when stored sample count >= windowSize; reset=TRUE clears it; invalid window clears it; recomputed every valid scan.
error/status: error=TRUE and status=16#8200 only when windowSize<1 or >100; otherwise FALSE/16#0000 (PUB004, PUB006, PUB007).
capture_priority: reset=TRUE suppresses capture; cyclicExecution=TRUE captures every scan and trigger has no effect; trigger uses one rising edge when cyclicExecution=FALSE.
window_resize: if a valid windowSize is smaller than stored count, oldest samples are discarded to the new width before capture; this detail is unspecified by PUB and implemented consistently.
boundaries: windowSize 1..100, circular buffer capacity 100 LREAL; divisor INT_TO_LREAL(local_count); windowSizeReached includes the equal boundary.
*)
(* CONTRACT_RULES [] *)

FUNCTION_BLOCK FB
VAR_INPUT
    cyclicExecution : BOOL;
    trigger : BOOL;
    value : LREAL;
    windowSize : INT;
    reset : BOOL;
END_VAR
VAR_OUTPUT
    average : LREAL;
    windowSizeReached : BOOL;
    error : BOOL;
    status : WORD;
END_VAR
VAR
    local_buffer : ARRAY[0..99] OF LREAL;
    local_count : INT := 0;
    local_head : INT := 0;
    local_sum : LREAL := 0.0;
    local_trigger_rt : R_TRIG;
    local_append_index : INT;
END_VAR

local_trigger_rt(CLK := trigger);

IF reset THEN
    local_count := 0;
    local_head := 0;
    local_sum := 0.0;
    average := 0.0;
    windowSizeReached := FALSE;
END_IF;

IF (windowSize < 1) OR (windowSize > 100) THEN
    error := TRUE;
    status := 16#8200;
    windowSizeReached := FALSE;
ELSE
    error := FALSE;
    status := 16#0000;

    WHILE local_count > windowSize DO
        local_sum := local_sum - local_buffer[local_head];
        local_head := (local_head + 1) MOD 100;
        local_count := local_count - 1;
    END_WHILE;

    IF local_count > 0 THEN
        average := local_sum / INT_TO_LREAL(local_count);
    ELSE
        average := 0.0;
    END_IF;

    windowSizeReached := local_count >= windowSize;

    IF NOT reset THEN
        IF cyclicExecution OR local_trigger_rt.Q THEN
            IF local_count < windowSize THEN
                local_append_index := (local_head + local_count) MOD 100;
                local_buffer[local_append_index] := value;
                local_sum := local_sum + value;
                local_count := local_count + 1;
            ELSE
                local_sum := local_sum - local_buffer[local_head] + value;
                local_buffer[local_head] := value;
                local_head := (local_head + 1) MOD 100;
            END_IF;

            IF local_count > 0 THEN
                average := local_sum / INT_TO_LREAL(local_count);
            END_IF;

            windowSizeReached := local_count >= windowSize;
        END_IF;
    END_IF;
END_IF;

END_FUNCTION_BLOCK

(* ---- public-medium-03.candidate_03.st ---- *)
(* ENGINEERING_CONTRACT
average: activates when a sample is accepted or the valid window changes; holds the last valid result otherwise; reset sets it to 0.0.
windowSizeReached: TRUE while retained sample count >= windowSize; reset or invalid window forces FALSE.
error/status: windowSize < 1 or windowSize > 100 sets error=TRUE and status=16#8200; a valid window sets error=FALSE and status=16#0000.
capture priority: cyclicExecution=TRUE captures every scan and suppresses trigger; trigger uses R_TRIG only while cyclicExecution=FALSE; reset suppresses capture.
window resize: shrinking removes the oldest points so only the most recent windowSize values remain; growing preserves retained points and continues filling without resetting.
reset: level-triggered on reset=TRUE; clears head, count, sum, average, and windowSizeReached.
invalid window preserves retained data but prevents new samples and forces windowSizeReached=FALSE.
Boundaries: windowSize is 1..100; storage is ARRAY[0..99] OF LREAL; average divides by INT_TO_LREAL(count).
PUB001, PUB002, PUB003, PUB004, PUB006, PUB007.
*)
(* CONTRACT_RULES [] *)

FUNCTION_BLOCK FB
VAR_INPUT
    cyclicExecution : BOOL;
    trigger : BOOL;
    value : LREAL;
    windowSize : INT;
    reset : BOOL;
END_VAR
VAR_OUTPUT
    average : LREAL;
    windowSizeReached : BOOL;
    error : BOOL;
    status : WORD;
END_VAR
VAR
    local_buffer : ARRAY[0..99] OF LREAL;
    local_count : INT;
    local_head : INT;
    local_sum : LREAL;
    local_to_remove : INT;
    local_insert_index : INT;
    local_trigger_rt : R_TRIG;
END_VAR

local_trigger_rt(CLK := trigger);

IF reset THEN
    local_count := 0;
    local_head := 0;
    local_sum := 0.0;
    average := 0.0;
    windowSizeReached := FALSE;
END_IF;

IF (windowSize < 1) OR (windowSize > 100) THEN
    error := TRUE;
    status := 16#8200;
    windowSizeReached := FALSE;
ELSE
    error := FALSE;
    status := 16#0000;

    IF local_count > windowSize THEN
        local_to_remove := local_count - windowSize;
        WHILE local_to_remove > 0 DO
            local_sum := local_sum - local_buffer[local_head];
            local_head := local_head + 1;
            IF local_head >= 100 THEN
                local_head := 0;
            END_IF;
            local_to_remove := local_to_remove - 1;
        END_WHILE;
        local_count := windowSize;
    END_IF;

    IF NOT reset THEN
        IF cyclicExecution OR (local_trigger_rt.Q AND (NOT cyclicExecution)) THEN
            IF local_count < windowSize THEN
                local_insert_index := (local_head + local_count) MOD 100;
                local_buffer[local_insert_index] := value;
                local_sum := local_sum + value;
                local_count := local_count + 1;
            ELSE
                local_sum := local_sum - local_buffer[local_head] + value;
                local_buffer[local_head] := value;
                local_head := local_head + 1;
                IF local_head >= 100 THEN
                    local_head := 0;
                END_IF;
            END_IF;
        END_IF;
    END_IF;

    IF local_count > 0 THEN
        average := local_sum / INT_TO_LREAL(local_count);
    END_IF;

    windowSizeReached := local_count >= windowSize;
END_IF;

END_FUNCTION_BLOCK

(* ---- public-medium-03.candidate_04.st ---- *)
(* ENGINEERING_CONTRACT
average: updated on each accepted sample; otherwise holds last valid result; reset sets it to 0.0; units/value domain follow input value (LREAL).
windowSizeReached: TRUE while retained sample count >= current valid windowSize; reset clears it; invalid window forces FALSE.
error/status: windowSize 1..100 -> FALSE/16#0000; otherwise -> TRUE/16#8200. Reset is evaluated before window validation.
capture priority: cyclicExecution=TRUE captures every scan and ignores trigger; otherwise R_TRIG trigger captures; reset suppresses capture in the same scan.
resize: a valid windowSize reduction shrinks retained history to the latest windowSize samples and recomputes average before capture.
PUB001, PUB002, PUB003, PUB004, PUB006, PUB007.
*)
(* CONTRACT_RULES [] *)

FUNCTION_BLOCK FB
VAR_INPUT
    cyclicExecution : BOOL;
    trigger : BOOL;
    value : LREAL;
    windowSize : INT;
    reset : BOOL;
END_VAR
VAR_OUTPUT
    average : LREAL;
    windowSizeReached : BOOL;
    error : BOOL;
    status : WORD;
END_VAR
VAR
    local_buffer : ARRAY[0..99] OF LREAL;
    local_count : INT;
    local_sum : LREAL;
    local_trigger_rt : R_TRIG;
    tmp_i : INT;
    tmp_old : LREAL;
END_VAR

local_trigger_rt(CLK := trigger);

IF reset THEN
    local_count := 0;
    local_sum := 0.0;
    average := 0.0;
    windowSizeReached := FALSE;
END_IF;

IF (windowSize < 1) OR (windowSize > 100) THEN
    error := TRUE;
    status := 16#8200;
    windowSizeReached := FALSE;
ELSE
    error := FALSE;
    status := 16#0000;

    WHILE local_count > windowSize DO
        local_sum := local_sum - local_buffer[0];
        IF local_count > 1 THEN
            FOR tmp_i := 0 TO local_count - 2 DO
                local_buffer[tmp_i] := local_buffer[tmp_i + 1];
            END_FOR;
        END_IF;
        local_count := local_count - 1;
    END_WHILE;

    IF local_count > 0 THEN
        average := local_sum / INT_TO_LREAL(local_count);
    END_IF;

    windowSizeReached := local_count >= windowSize;

    IF NOT reset THEN
        IF cyclicExecution OR local_trigger_rt.Q THEN
            IF local_count < windowSize THEN
                local_buffer[local_count] := value;
                local_sum := local_sum + value;
                local_count := local_count + 1;
            ELSE
                tmp_old := local_buffer[0];
                IF local_count > 1 THEN
                    FOR tmp_i := 0 TO local_count - 2 DO
                        local_buffer[tmp_i] := local_buffer[tmp_i + 1];
                    END_FOR;
                END_IF;
                local_buffer[local_count - 1] := value;
                local_sum := local_sum - tmp_old + value;
            END_IF;

            IF local_count > 0 THEN
                average := local_sum / INT_TO_LREAL(local_count);
            END_IF;

            windowSizeReached := local_count >= windowSize;
        END_IF;
    END_IF;
END_IF;

END_FUNCTION_BLOCK

(* ---- public-medium-03.raw_candidate_01.st ---- *)
(* ENGINEERING_CONTRACT
average: activated when a sample is accepted; otherwise holds last valid result; reset sets it to 0.0; units are inherited from value (LREAL).
windowSizeReached: TRUE when accepted sample count >= windowSize; holds until reset or invalid window; no edge-only behavior.
error/status: windowSize < 1 or windowSize > 100 sets error=TRUE and status=16#8200; valid window sets error=FALSE and status=16#0000.
capture priority: cyclicExecution=TRUE captures every scan and suppresses trigger; trigger uses R_TRIG only while cyclicExecution=FALSE; reset suppresses capture.
reset: level-triggered on reset=TRUE, clears sum, buffer count, write index, average, and windowSizeReached.
invalid window preserves accumulated average data but forces windowSizeReached=FALSE and prevents new samples.
Boundaries: windowSize is 1..100; storage is ARRAY[0..99] OF LREAL; average division uses INT_TO_LREAL.
PUB001, PUB002, PUB003, PUB004, PUB006, PUB007.
*)
(* CONTRACT_RULES [] *)

FUNCTION_BLOCK FB
VAR_INPUT
    cyclicExecution : BOOL;
    trigger : BOOL;
    value : LREAL;
    windowSize : INT;
    reset : BOOL;
END_VAR
VAR_OUTPUT
    average : LREAL;
    windowSizeReached : BOOL;
    error : BOOL;
    status : WORD;
END_VAR
VAR
    local_buffer : ARRAY[0..99] OF LREAL;
    local_count : INT;
    local_write_index : INT;
    local_sum : LREAL;
    local_trigger_rt : R_TRIG;
END_VAR

local_trigger_rt(CLK := trigger);

IF reset THEN
    local_count := 0;
    local_write_index := 0;
    local_sum := 0.0;
    average := 0.0;
    windowSizeReached := FALSE;
END_IF;

IF (windowSize < 1) OR (windowSize > 100) THEN
    error := TRUE;
    status := 16#8200;
    windowSizeReached := FALSE;
ELSE
    error := FALSE;
    status := 16#0000;

    IF NOT reset THEN
        IF cyclicExecution OR (local_trigger_rt.Q AND (NOT cyclicExecution)) THEN
            IF local_count < windowSize THEN
                local_buffer[local_count] := value;
                local_sum := local_sum + value;
                local_count := local_count + 1;
            ELSE
                local_sum := local_sum - local_buffer[local_write_index] + value;
                local_buffer[local_write_index] := value;
                local_write_index := local_write_index + 1;
                IF local_write_index >= windowSize THEN
                    local_write_index := 0;
                END_IF;
            END_IF;

            IF local_count > 0 THEN
                average := local_sum / INT_TO_LREAL(local_count);
            END_IF;

            windowSizeReached := local_count >= windowSize;
        END_IF;
    END_IF;
END_IF;

END_FUNCTION_BLOCK

(* ---- public-medium-03.raw_candidate_02.st ---- *)
(* ENGINEERING_CONTRACT
average: updates on each accepted sample (PUB002/PUB003), holds between samples; reset=TRUE clears it in the same scan; units LREAL.
windowSizeReached: TRUE when stored sample count >= windowSize; reset=TRUE clears it; invalid window clears it; recomputed every valid scan.
error/status: error=TRUE and status=16#8200 only when windowSize<1 or >100; otherwise FALSE/16#0000 (PUB004, PUB006, PUB007).
capture_priority: reset=TRUE suppresses capture; cyclicExecution=TRUE captures every scan and trigger has no effect; trigger uses one rising edge when cyclicExecution=FALSE.
window_resize: if a valid windowSize is smaller than stored count, oldest samples are discarded to the new width before capture; this detail is unspecified by PUB and implemented consistently.
boundaries: windowSize 1..100, circular buffer capacity 100 LREAL; divisor INT_TO_LREAL(local_count); windowSizeReached includes the equal boundary.
*)
(* CONTRACT_RULES [] *)

FUNCTION_BLOCK FB
VAR_INPUT
    cyclicExecution : BOOL;
    trigger : BOOL;
    value : LREAL;
    windowSize : INT;
    reset : BOOL;
END_VAR
VAR_OUTPUT
    average : LREAL;
    windowSizeReached : BOOL;
    error : BOOL;
    status : WORD;
END_VAR
VAR
    local_buffer : ARRAY[0..99] OF LREAL;
    local_count : INT := 0;
    local_head : INT := 0;
    local_sum : LREAL := 0.0;
    local_trigger_rt : R_TRIG;
    local_append_index : INT;
END_VAR

local_trigger_rt(CLK := trigger);

IF reset THEN
    local_count := 0;
    local_head := 0;
    local_sum := 0.0;
    average := 0.0;
    windowSizeReached := FALSE;
END_IF;

IF (windowSize < 1) OR (windowSize > 100) THEN
    error := TRUE;
    status := 16#8200;
    windowSizeReached := FALSE;
ELSE
    error := FALSE;
    status := 16#0000;

    WHILE local_count > windowSize DO
        local_sum := local_sum - local_buffer[local_head];
        local_head := (local_head + 1) MOD 100;
        local_count := local_count - 1;
    END_WHILE;

    IF local_count > 0 THEN
        average := local_sum / INT_TO_LREAL(local_count);
    ELSE
        average := 0.0;
    END_IF;

    windowSizeReached := local_count >= windowSize;

    IF NOT reset THEN
        IF cyclicExecution OR local_trigger_rt.Q THEN
            IF local_count < windowSize THEN
                local_append_index := (local_head + local_count) MOD 100;
                local_buffer[local_append_index] := value;
                local_sum := local_sum + value;
                local_count := local_count + 1;
            ELSE
                local_sum := local_sum - local_buffer[local_head] + value;
                local_buffer[local_head] := value;
                local_head := (local_head + 1) MOD 100;
            END_IF;

            IF local_count > 0 THEN
                average := local_sum / INT_TO_LREAL(local_count);
            END_IF;

            windowSizeReached := local_count >= windowSize;
        END_IF;
    END_IF;
END_IF;

END_FUNCTION_BLOCK

(* ---- public-medium-03.raw_candidate_03.st ---- *)
(* ENGINEERING_CONTRACT
average: activates when a sample is accepted or the valid window changes; holds the last valid result otherwise; reset sets it to 0.0.
windowSizeReached: TRUE while retained sample count >= windowSize; reset or invalid window forces FALSE.
error/status: windowSize < 1 or windowSize > 100 sets error=TRUE and status=16#8200; a valid window sets error=FALSE and status=16#0000.
capture priority: cyclicExecution=TRUE captures every scan and suppresses trigger; trigger uses R_TRIG only while cyclicExecution=FALSE; reset suppresses capture.
window resize: shrinking removes the oldest points so only the most recent windowSize values remain; growing preserves retained points and continues filling without resetting.
reset: level-triggered on reset=TRUE; clears head, count, sum, average, and windowSizeReached.
invalid window preserves retained data but prevents new samples and forces windowSizeReached=FALSE.
Boundaries: windowSize is 1..100; storage is ARRAY[0..99] OF LREAL; average divides by INT_TO_LREAL(count).
PUB001, PUB002, PUB003, PUB004, PUB006, PUB007.
*)
(* CONTRACT_RULES [] *)

FUNCTION_BLOCK FB
VAR_INPUT
    cyclicExecution : BOOL;
    trigger : BOOL;
    value : LREAL;
    windowSize : INT;
    reset : BOOL;
END_VAR
VAR_OUTPUT
    average : LREAL;
    windowSizeReached : BOOL;
    error : BOOL;
    status : WORD;
END_VAR
VAR
    local_buffer : ARRAY[0..99] OF LREAL;
    local_count : INT;
    local_head : INT;
    local_sum : LREAL;
    local_to_remove : INT;
    local_insert_index : INT;
    local_trigger_rt : R_TRIG;
END_VAR

local_trigger_rt(CLK := trigger);

IF reset THEN
    local_count := 0;
    local_head := 0;
    local_sum := 0.0;
    average := 0.0;
    windowSizeReached := FALSE;
END_IF;

IF (windowSize < 1) OR (windowSize > 100) THEN
    error := TRUE;
    status := 16#8200;
    windowSizeReached := FALSE;
ELSE
    error := FALSE;
    status := 16#0000;

    IF local_count > windowSize THEN
        local_to_remove := local_count - windowSize;
        WHILE local_to_remove > 0 DO
            local_sum := local_sum - local_buffer[local_head];
            local_head := local_head + 1;
            IF local_head >= 100 THEN
                local_head := 0;
            END_IF;
            local_to_remove := local_to_remove - 1;
        END_WHILE;
        local_count := windowSize;
    END_IF;

    IF NOT reset THEN
        IF cyclicExecution OR (local_trigger_rt.Q AND (NOT cyclicExecution)) THEN
            IF local_count < windowSize THEN
                local_insert_index := (local_head + local_count) MOD 100;
                local_buffer[local_insert_index] := value;
                local_sum := local_sum + value;
                local_count := local_count + 1;
            ELSE
                local_sum := local_sum - local_buffer[local_head] + value;
                local_buffer[local_head] := value;
                local_head := local_head + 1;
                IF local_head >= 100 THEN
                    local_head := 0;
                END_IF;
            END_IF;
        END_IF;
    END_IF;

    IF local_count > 0 THEN
        average := local_sum / INT_TO_LREAL(local_count);
    END_IF;

    windowSizeReached := local_count >= windowSize;
END_IF;

END_FUNCTION_BLOCK

(* ---- public-medium-03.raw_candidate_04.st ---- *)
(* ENGINEERING_CONTRACT
average: updated on each accepted sample; otherwise holds last valid result; reset sets it to 0.0; units/value domain follow input value (LREAL).
windowSizeReached: TRUE while retained sample count >= current valid windowSize; reset clears it; invalid window forces FALSE.
error/status: windowSize 1..100 -> FALSE/16#0000; otherwise -> TRUE/16#8200. Reset is evaluated before window validation.
capture priority: cyclicExecution=TRUE captures every scan and ignores trigger; otherwise R_TRIG trigger captures; reset suppresses capture in the same scan.
resize: a valid windowSize reduction shrinks retained history to the latest windowSize samples and recomputes average before capture.
PUB001, PUB002, PUB003, PUB004, PUB006, PUB007.
*)
(* CONTRACT_RULES [] *)

FUNCTION_BLOCK FB
VAR_INPUT
    cyclicExecution : BOOL;
    trigger : BOOL;
    value : LREAL;
    windowSize : INT;
    reset : BOOL;
END_VAR
VAR_OUTPUT
    average : LREAL;
    windowSizeReached : BOOL;
    error : BOOL;
    status : WORD;
END_VAR
VAR
    local_buffer : ARRAY[0..99] OF LREAL;
    local_count : INT;
    local_sum : LREAL;
    local_trigger_rt : R_TRIG;
    tmp_i : INT;
    tmp_old : LREAL;
END_VAR

local_trigger_rt(CLK := trigger);

IF reset THEN
    local_count := 0;
    local_sum := 0.0;
    average := 0.0;
    windowSizeReached := FALSE;
END_IF;

IF (windowSize < 1) OR (windowSize > 100) THEN
    error := TRUE;
    status := 16#8200;
    windowSizeReached := FALSE;
ELSE
    error := FALSE;
    status := 16#0000;

    WHILE local_count > windowSize DO
        local_sum := local_sum - local_buffer[0];
        IF local_count > 1 THEN
            FOR tmp_i := 0 TO local_count - 2 DO
                local_buffer[tmp_i] := local_buffer[tmp_i + 1];
            END_FOR;
        END_IF;
        local_count := local_count - 1;
    END_WHILE;

    IF local_count > 0 THEN
        average := local_sum / INT_TO_LREAL(local_count);
    END_IF;

    windowSizeReached := local_count >= windowSize;

    IF NOT reset THEN
        IF cyclicExecution OR local_trigger_rt.Q THEN
            IF local_count < windowSize THEN
                local_buffer[local_count] := value;
                local_sum := local_sum + value;
                local_count := local_count + 1;
            ELSE
                tmp_old := local_buffer[0];
                IF local_count > 1 THEN
                    FOR tmp_i := 0 TO local_count - 2 DO
                        local_buffer[tmp_i] := local_buffer[tmp_i + 1];
                    END_FOR;
                END_IF;
                local_buffer[local_count - 1] := value;
                local_sum := local_sum - tmp_old + value;
            END_IF;

            IF local_count > 0 THEN
                average := local_sum / INT_TO_LREAL(local_count);
            END_IF;

            windowSizeReached := local_count >= windowSize;
        END_IF;
    END_IF;
END_IF;

END_FUNCTION_BLOCK

(* ---- public-medium-04.candidate_01.st ---- *)
FUNCTION_BLOCK FB
VAR_INPUT
    TemperatureSensorInput : REAL;
    SetTemperature : REAL;
END_VAR
VAR_OUTPUT
    CurrentTemperature : REAL;
    SetTempDisplay : REAL;
    HeaterStatus : BOOL;
    OverheatProtection : BOOL;
    HeaterOutput : BOOL;
END_VAR
VAR
    local_SensorFault : BOOL;
    local_HeatCommand : BOOL;
    local_OverheatActive : BOOL;
    HeaterContinuousTimer : TON;
    OverheatCooldownTimer : TON;
END_VAR

(*
ENGINEERING_CONTRACT
- Displays follow inputs each scan; REAL preserved without conversion (PUB002/PUB007).
- Normal heat: on when TemperatureSensorInput < SetTemperature; off when >= SetTemperature.
  Equality is unspecified by PUB003-PUB005 and is interpreted as off.
- Sensor fault: TemperatureSensorInput < 0.0 OR TemperatureSensorInput > 100.0 forces heat off.
  Values 0.0 and 100.0 remain valid (PUB008).
- Overheat: continuous HeaterOutput TRUE for 5 s starts protection; heater is forced off and
  OverheatProtection stays TRUE for a 3 s cooldown, then clears automatically (PUB006).
- Same-scan priority: sensor fault / active overheat overrides normal demand; a 5 s timer hit
  overrides the computed heat command in that scan.
- Units/boundaries: TIME uses T#5S and T#3S.
*)
(* CONTRACT_RULES [] *)

CurrentTemperature := TemperatureSensorInput;
SetTempDisplay := SetTemperature;

local_SensorFault := (TemperatureSensorInput < 0.0) OR (TemperatureSensorInput > 100.0);

IF local_OverheatActive THEN
    OverheatCooldownTimer(IN := TRUE, PT := T#3S);
    IF OverheatCooldownTimer.Q THEN
        local_OverheatActive := FALSE;
    END_IF;
ELSE
    OverheatCooldownTimer(IN := FALSE, PT := T#3S);
END_IF;

IF local_SensorFault OR local_OverheatActive THEN
    local_HeatCommand := FALSE;
ELSIF TemperatureSensorInput < SetTemperature THEN
    local_HeatCommand := TRUE;
ELSE
    local_HeatCommand := FALSE;
END_IF;

HeaterContinuousTimer(IN := local_HeatCommand, PT := T#5S);
IF HeaterContinuousTimer.Q THEN
    local_OverheatActive := TRUE;
    local_HeatCommand := FALSE;
END_IF;

HeaterOutput := local_HeatCommand AND NOT local_SensorFault AND NOT local_OverheatActive;
HeaterStatus := HeaterOutput;
OverheatProtection := local_OverheatActive;

END_FUNCTION_BLOCK

(* ---- public-medium-04.candidate_02.st ---- *)
FUNCTION_BLOCK FB
VAR_INPUT
    TemperatureSensorInput : REAL;
    SetTemperature : REAL;
END_VAR
VAR_OUTPUT
    CurrentTemperature : REAL;
    SetTempDisplay : REAL;
    HeaterStatus : BOOL;
    OverheatProtection : BOOL;
    HeaterOutput : BOOL;
END_VAR
VAR
    local_SensorFault : BOOL;
    local_HeatCommand : BOOL;
    local_OverheatActive : BOOL;
    HeaterContinuousTimer : TON;
    OverheatCooldownTimer : TON;
END_VAR

(*
ENGINEERING_CONTRACT
- Displays follow inputs each scan; REAL values are passed through without conversion (PUB002/PUB007).
- Normal heat: on when TemperatureSensorInput < SetTemperature; off when TemperatureSensorInput >= SetTemperature.
  Equality is unspecified by PUB003-PUB005 and is interpreted as off.
- Sensor fault: TemperatureSensorInput < 0.0 OR TemperatureSensorInput > 100.0 forces heat off.
  Values 0.0 and 100.0 remain valid (PUB008).
- Overheat: triggered only after continuous heating exceeds 5 s (strict > boundary implemented as
  T#5001MS). The trip starts a 3 s release timer; HeaterOutput remains off and OverheatProtection
  clears when the release timer reaches T#3S (PUB006).
- Same-scan priority: sensor fault / active overheat overrides normal demand; a continuous-heat
  timer trip overrides the computed heat command in that scan and starts the release timer.
- Units/boundaries: TIME uses T#5001MS for the heat trip and T#3S for release.
*)

(* CONTRACT_RULES [] *)

CurrentTemperature := TemperatureSensorInput;
SetTempDisplay := SetTemperature;

local_SensorFault := (TemperatureSensorInput < 0.0) OR (TemperatureSensorInput > 100.0);

IF local_SensorFault OR local_OverheatActive THEN
    local_HeatCommand := FALSE;
ELSIF TemperatureSensorInput < SetTemperature THEN
    local_HeatCommand := TRUE;
ELSE
    local_HeatCommand := FALSE;
END_IF;

HeaterContinuousTimer(IN := local_HeatCommand, PT := T#5001MS);
IF HeaterContinuousTimer.Q THEN
    local_OverheatActive := TRUE;
    local_HeatCommand := FALSE;
END_IF;

IF local_OverheatActive THEN
    OverheatCooldownTimer(IN := TRUE, PT := T#3S);
    IF OverheatCooldownTimer.Q THEN
        local_OverheatActive := FALSE;
    END_IF;
ELSE
    OverheatCooldownTimer(IN := FALSE, PT := T#3S);
END_IF;

HeaterOutput := local_HeatCommand AND NOT local_SensorFault AND NOT local_OverheatActive;
HeaterStatus := HeaterOutput;
OverheatProtection := local_OverheatActive;

END_FUNCTION_BLOCK

(* ---- public-medium-04.raw_candidate_01.st ---- *)
FUNCTION_BLOCK FB
VAR_INPUT
    TemperatureSensorInput : REAL;
    SetTemperature : REAL;
END_VAR
VAR_OUTPUT
    CurrentTemperature : REAL;
    SetTempDisplay : REAL;
    HeaterStatus : BOOL;
    OverheatProtection : BOOL;
    HeaterOutput : BOOL;
END_VAR
VAR
    local_SensorFault : BOOL;
    local_HeatCommand : BOOL;
    local_OverheatActive : BOOL;
    HeaterContinuousTimer : TON;
    OverheatCooldownTimer : TON;
END_VAR

(*
ENGINEERING_CONTRACT
- Displays follow inputs each scan; REAL preserved without conversion (PUB002/PUB007).
- Normal heat: on when TemperatureSensorInput < SetTemperature; off when >= SetTemperature.
  Equality is unspecified by PUB003-PUB005 and is interpreted as off.
- Sensor fault: TemperatureSensorInput < 0.0 OR TemperatureSensorInput > 100.0 forces heat off.
  Values 0.0 and 100.0 remain valid (PUB008).
- Overheat: continuous HeaterOutput TRUE for 5 s starts protection; heater is forced off and
  OverheatProtection stays TRUE for a 3 s cooldown, then clears automatically (PUB006).
- Same-scan priority: sensor fault / active overheat overrides normal demand; a 5 s timer hit
  overrides the computed heat command in that scan.
- Units/boundaries: TIME uses T#5S and T#3S.
*)
(* CONTRACT_RULES [] *)

CurrentTemperature := TemperatureSensorInput;
SetTempDisplay := SetTemperature;

local_SensorFault := (TemperatureSensorInput < 0.0) OR (TemperatureSensorInput > 100.0);

IF local_OverheatActive THEN
    OverheatCooldownTimer(IN := TRUE, PT := T#3S);
    IF OverheatCooldownTimer.Q THEN
        local_OverheatActive := FALSE;
    END_IF;
ELSE
    OverheatCooldownTimer(IN := FALSE, PT := T#3S);
END_IF;

IF local_SensorFault OR local_OverheatActive THEN
    local_HeatCommand := FALSE;
ELSIF TemperatureSensorInput < SetTemperature THEN
    local_HeatCommand := TRUE;
ELSE
    local_HeatCommand := FALSE;
END_IF;

HeaterContinuousTimer(IN := local_HeatCommand, PT := T#5S);
IF HeaterContinuousTimer.Q THEN
    local_OverheatActive := TRUE;
    local_HeatCommand := FALSE;
END_IF;

HeaterOutput := local_HeatCommand AND NOT local_SensorFault AND NOT local_OverheatActive;
HeaterStatus := HeaterOutput;
OverheatProtection := local_OverheatActive;

END_FUNCTION_BLOCK
